(* IEC 61131-3 sources: JingjiangArm/moonboxpro_arm_8.4/Application/Application/任务列表/TensionTask/电机运动/MotionCtl_Gear, 17 files *)

(* ---- StMotorParam_Vel.st ---- *)
(*@CES
Name=StMotorParam_Vel
Type=Gvl
TypeGuid=2db5746d-d284-4425-9f7f-2663a34b0ebc
Guid=35fd48d6-a97b-4a50-89b7-bfdefdaf1e25
HasDeclaration=True
HasImplementation=False
*)
{DECLARATION}
TYPE StMotorParam_Vel :(*速度运动同步轴就是这些各参数了*)
STRUCT
	iAxisId: INT;
	iCoreId: INT;
	iStationId: INT;
	iMoveStep: INT;
	iMotionMode: INT;(*运动模式-=0：电子齿轮=1：JOG=2：点位*)
	xMoveRev: BOOL;
	xMoveEn: BOOL;
	rAxisGirth: REAL;(*同步版周*)
	xMoveVelMode: BOOL;(*=0:线速度=1转速*)
	rAxisVel: REAL;(*速度*)
	uiAxisNum: UINT;(*减速比分子*)
	uiAxisDen: UINT;(*减速比分母*)
	liTargetPos: LINT;(*点位目标位置*)
	udiTargetVel: UDINT;

	//2026.01.31.130843 | + | 增加停机维持伺服功能 秦华有停机维持伺服的功能，需要增加一个判断是否是使能状态的标志
	xAxisOn_ing : BOOL;//此标志表示该轴正处于使能中。。。

	//2026.05.09.085650 | + | 将大指令写入的值先放在这里，然后再穿进去
	modify_delta: DINT;
	/// 可以为正值
	ratio_a: DINT;
	/// 必须为正值
	ratio_b: DINT;

	//2026.05.12.201038 | + | 增加轴单运行中的标志
	xAxisInching : BOOL;
END_STRUCT
END_TYPE

{IMPLEMENTATION}

(* ---- KS_SetMotionCheckServoOn.st ---- *)
(*@CES
Name=KS_SetMotionCheckServoOn
Type=FunctionBlock
TypeGuid=6f9dac99-8de1-4efc-8465-68ac443b7d08
Guid=16f739cf-935e-4f65-a185-0fbe09498330
HasDeclaration=True
HasImplementation=True
*)
{DECLARATION}
FUNCTION KS_SetMotionCheckServoOn : INT
VAR_INPUT
	i_iAxisId: INT;
	i_iCoreId: INT;
	i_iStationId: INT;
	i_pxMoveEn : POINTER TO BOOL;
	i_dwMotionSts: DWORD;
	i_dwDriverSts: DWORD;
	i_pxServoOn: POINTER TO BOOL;
	i_pstStHYLogFifo			: POINTER TO StHYLogFifo;(* 2025.8.23.170701/han.dp/增加的日志队列 *)
END_VAR
VAR
	iResult: INT;
	xRtn: BOOL;
	iFailedAxisCntNum: INT;
	wLogLevel: WORD;
	sMsg_major: STRING;
	sMsg_minor: STRING;
END_VAR

{IMPLEMENTATION}
iResult:= 0;
sMsg_major:= ''; (* 2021.2.26.170203/ *)
sMsg_minor:= ''; (* 2021.2.26.170203/ *)
IF i_iStationId>=1 AND i_iStationId<=MAX_STATION_NUM AND
	i_iAxisId>=1 AND i_iAxisId<=MAX_STATION_NUM AND
	(i_iCoreId=1 OR i_iCoreId=2) THEN

	IF i_pxServoOn^ AND i_pxMoveEn^ THEN
		xRtn:= (*i_dwDriverSts.1 AND*) i_dwMotionSts.9;

		IF NOT xRtn THEN
			iResult:= iResult+1;
			(* 2021.2.26.172210/归属于普通报警 *)
			wLogLevel:= LOG_LEVEL_ALARM_NORMAL;
	(*2022.6.4.093146|精简打印信息！*)
	(*		sMsg_major:= CONCAT('ALARM_NORMAL: KS_SetGrpAxisClrSts_PshLog|Aid:', INT_TO_STRING(iAxisId));*)
			sMsg_major:= CONCAT('KS_SetMotionCheckServoOn|Aid:', INT_TO_STRING(i_iAxisId));
			sMsg_major:= CONCAT(sMsg_major, '|Sid:');
			sMsg_major:= CONCAT(sMsg_major, INT_TO_STRING(i_iStationId));
			sMsg_minor:= CONCAT('CheckServoOn|', BOOL_TO_STRING(xRtn));
			sMsg_minor:= CONCAT(sMsg_minor,'|MotionSts:');
			sMsg_minor:= CONCAT(sMsg_minor, DWORD_TO_STRING(i_dwMotionSts));
		END_IF

		//i_pxServoOn^:= FALSE;
	END_IF
END_IF

IF sMsg_major<>'' THEN (* 2021.2.26.172055/有内容代表要写日志的 *)
	KS_HY_AddMsgToLog(i_pstStHYLogFifo, wLogLevel, sMsg_major, sMsg_minor);
END_IF

KS_SetMotionCheckServoOn:= iResult;

(* ---- KS_SetMotionClrSts.st ---- *)
(*@CES
Name=KS_SetMotionClrSts
Type=FunctionBlock
TypeGuid=6f9dac99-8de1-4efc-8465-68ac443b7d08
Guid=5963aa42-d132-45f6-9961-fbcc83163ad5
HasDeclaration=True
HasImplementation=True
*)
{DECLARATION}
FUNCTION KS_SetMotionClrSts : INT(*0:无错误| >0:失败的指令数量; |-1:参数错误;*)
VAR_INPUT
	i_iAxisId: INT;
	i_iCoreId: INT;
	i_iStationId: INT;
	i_pstStHYLogFifo			: POINTER TO StHYLogFifo;(* 2025.8.23.170701/han.dp/增加的日志队列 *)
END_VAR
VAR
	iResult: INT;
	iRtn: INT;
	iFailedAxisCntNum: INT;
	wLogLevel: WORD;
	sMsg_major: STRING;
	sMsg_minor: STRING;
END_VAR

{IMPLEMENTATION}
iResult:= 0;
sMsg_major:= ''; (* 2021.2.26.170203/ *)
sMsg_minor:= ''; (* 2021.2.26.170203/ *)
IF i_iStationId>=1 AND i_iStationId<=MAX_STATION_NUM AND
	i_iAxisId>=1 AND i_iAxisId<=MAX_STATION_NUM AND
	(i_iCoreId=1 OR i_iCoreId=2) THEN
	iRtn:= GTN_ClrSts(i_iCoreId, i_iAxisId, 1);(*清除错误|*)
	IF iRtn<>0 THEN
		iResult:= iRtn;
		(* 2021.2.26.172210/归属于普通报警 *)
		wLogLevel:= LOG_LEVEL_ALARM;
(*2022.6.4.093146|精简打印信息！*)
(*		sMsg_major:= CONCAT('ALARM_NORMAL: KS_SetGrpAxisClrSts_PshLog|Aid:', INT_TO_STRING(iAxisId));*)
		sMsg_major:= CONCAT('KS_SetMotionClrSts|Aid:', INT_TO_STRING(i_iAxisId));
		sMsg_major:= CONCAT(sMsg_major, '|Sid:');
		sMsg_major:= CONCAT(sMsg_major, INT_TO_STRING(i_iStationId));
		sMsg_minor:= CONCAT('GTN_ClrSts: ', INT_TO_STRING(iRtn));
	END_IF
END_IF

IF sMsg_major<>'' THEN (* 2021.2.26.172055/有内容代表要写日志的 *)
	KS_HY_AddMsgToLog(i_pstStHYLogFifo, wLogLevel, sMsg_major, sMsg_minor);
END_IF

KS_SetMotionClrSts:= iResult;

(* ---- KS_SetMotionMode.st ---- *)
(*@CES
Name=KS_SetMotionMode
Type=FunctionBlock
TypeGuid=6f9dac99-8de1-4efc-8465-68ac443b7d08
Guid=eb1bfde3-c781-4a8b-bb4b-64a6f57a70ed
HasDeclaration=True
HasImplementation=True
*)
{DECLARATION}
FUNCTION KS_SetMotionMode : INT(*0:无错误| >0:失败的指令数量; |-1:参数错误;*)
VAR_INPUT
	i_iAxisId: INT;
	i_iCoreId: INT;
	i_iStationId: INT;
	i_iMoveMode: INT;
	i_iAxisId_Master: INT;
	i_xMasterType : BOOL;
	i_pstStHYLogFifo			: POINTER TO StHYLogFifo;(* 2025.8.23.170701/han.dp/增加的日志队列 *)
END_VAR
VAR
	iResult: INT;
	iRtn: INT;
	iFailedAxisCntNum: INT;
	wLogLevel: WORD;
	sMsg_major: STRING;
	sMsg_minor: STRING;
END_VAR

{IMPLEMENTATION}
iResult:= 0;
sMsg_major:= ''; (* 2021.2.26.170203/ *)
sMsg_minor:= ''; (* 2021.2.26.170203/ *)
IF i_iStationId>=1 AND i_iStationId<=MAX_STATION_NUM AND
	i_iAxisId>=1 AND i_iAxisId<=MAX_STATION_NUM AND
	(i_iCoreId=1 OR i_iCoreId=2) THEN
	IF i_iMoveMode=0 THEN
		iRtn := SetPrfGearModePrm(
				i_iCore:= i_iCoreId,
				i_iAxisId:= i_iAxisId,
				i_iMasterIndex:= i_iAxisId_Master,//i_pastTStGearParamUser^[iCnt_GearAxis].iMasterIndex,
				i_diMasterEven:= 1,//i_pastTStGearParamUser^[iCnt_GearAxis].diMasterEven,
				i_diSlaveEven:= 1,//i_pastTStGearParamUser^[iCnt_GearAxis].diSlaveEven,
				i_diMasterSlope:= 100000,
				i_xMasterType := i_xMasterType);//i_pastTStGearParamUser^[iCnt_GearAxis].diMasterSlope);

	ELSIF i_iMoveMode=1 THEN
		//2025.10.28.105106 | bai.zy  | 单运行仍然使用电子齿轮
		iRtn := SetPrfGearModePrm(
				i_iCore:= i_iCoreId,
				i_iAxisId:= i_iAxisId,
				i_iMasterIndex:= i_iAxisId_Master,//i_pastTStGearParamUser^[iCnt_GearAxis].iMasterIndex,
				i_diMasterEven:= 1,//i_pastTStGearParamUser^[iCnt_GearAxis].diMasterEven,
				i_diSlaveEven:= 1,//i_pastTStGearParamUser^[iCnt_GearAxis].diSlaveEven,
				i_diMasterSlope:= 100000,
				i_xMasterType := i_xMasterType);//i_pastTStGearParamUser^[iCnt_GearAxis].diMasterSlope);

// 		iRtn := SetPrfJogModePrm(
// 				i_iCore:= i_iCoreId,
// 				i_iAxisId:= i_iAxisId,
// 				i_lrAcc:= 1,
// 				i_lrDec:= 1,
// 				i_rSmooth:= 0.8);

	ELSIF i_iMoveMode=2 THEN
		iRtn := SetPrfTrapModePrm(
				i_iCoreId:= i_iCoreId,
				i_iAxisId:= i_iAxisId,
				i_lrVel:= 100,//i_pastTStTrapParamUser^[iCnt_TrapAxis].lrVel,
				i_lrAcc:= 2.0,//i_pastTStTrapParamUser^[iCnt_TrapAxis].lrAcc,
				i_lrDec:= 2.0,//i_pastTStTrapParamUser^[iCnt_TrapAxis].lrDec,
				i_iSmoothTime:= 0);//i_pastTStTrapParamUser^[iCnt_TrapAxis].iSmoothTime);
	ELSIF i_iMoveMode=3 THEN//增加一种运动模式2026.4.27.215724|收放料速度模式
		iRtn := SetPrfJogModePrm(
				i_iCore:= i_iCoreId,
				i_iAxisId:= i_iAxisId,
				i_lrAcc:= 1,
				i_lrDec:= 1,
				i_rSmooth:= 0.8);

	ELSE;
		iRtn := SetPrfGearModePrm(
				i_iCore:= i_iCoreId,
				i_iAxisId:= i_iAxisId,
				i_iMasterIndex:= i_iAxisId_Master,//i_pastTStGearParamUser^[iCnt_GearAxis].iMasterIndex,
				i_diMasterEven:= 1,//i_pastTStGearParamUser^[iCnt_GearAxis].diMasterEven,
				i_diSlaveEven:= 1,//i_pastTStGearParamUser^[iCnt_GearAxis].diSlaveEven,
				i_diMasterSlope:= 100000,
				i_xMasterType := i_xMasterType);//i_pastTStGearParamUser^[iCnt_GearAxis].diMasterSlope);
	END_IF

	IF iRtn<>0 THEN
		iResult:= iRtn;
		(* 2021.2.26.172210/归属于普通报警 *)
		wLogLevel:= LOG_LEVEL_ALARM;
(*2022.6.4.093146|精简打印信息！*)
(*		sMsg_major:= CONCAT('ALARM_NORMAL: KS_SetGrpAxisClrSts_PshLog|Aid:', INT_TO_STRING(iAxisId));*)
		sMsg_major:= CONCAT('KS_SetMotionMode|Aid:', INT_TO_STRING(i_iAxisId));
		sMsg_major:= CONCAT(sMsg_major, '|Sid:');
		sMsg_major:= CONCAT(sMsg_major, INT_TO_STRING(i_iStationId));
		//sMsg_minor:= CONCAT('GTN_ClrSts: ', INT_TO_STRING(iRtn));
	END_IF
END_IF

IF sMsg_major<>'' THEN (* 2021.2.26.172055/有内容代表要写日志的 *)
	KS_HY_AddMsgToLog(i_pstStHYLogFifo, wLogLevel, sMsg_major, sMsg_minor);
END_IF

KS_SetMotionMode:= iResult;

(* ---- KS_SetMotionServoOff.st ---- *)
(*@CES
Name=KS_SetMotionServoOff
Type=FunctionBlock
TypeGuid=6f9dac99-8de1-4efc-8465-68ac443b7d08
Guid=af78d755-d488-4f6e-8233-0470695debbc
HasDeclaration=True
HasImplementation=True
*)
{DECLARATION}
FUNCTION KS_SetMotionServoOff : INT(*0:无错误| >0:失败的指令数量; |-1:参数错误;*)
VAR_INPUT
	i_iAxisId: INT;
	i_iCoreId: INT;
	i_iStationId: INT;
	i_xForceAxisOff:BOOL;(*强制下伺服标志|有效后直接调用AXISOFF指令|2021.5.8.161449*)
	i_dwMotionSts: DWORD;
	i_dwDriverSts: DWORD;
	i_pxServoOn: POINTER TO BOOL;
	i_pstStHYLogFifo			: POINTER TO StHYLogFifo;(* 2025.8.23.170701/han.dp/增加的日志队列 *)
END_VAR
VAR
	iResult: INT;
	iRtn: INT;
	iFailedAxisCntNum: INT;
	wLogLevel: WORD;
	sMsg_major: STRING;
	sMsg_minor: STRING;
END_VAR

{IMPLEMENTATION}
iResult:= 0;
sMsg_major:= ''; (* 2021.2.26.170203/ *)
sMsg_minor:= ''; (* 2021.2.26.170203/ *)
IF i_iStationId>=1 AND i_iStationId<=MAX_STATION_NUM AND
	i_iAxisId>=1 AND i_iAxisId<=MAX_STATION_NUM AND
	(i_iCoreId=1 OR i_iCoreId=2) THEN

	IF i_pxServoOn^ (*OR i_dwDriverSts.1*) THEN
		IF i_xForceAxisOff THEN
			iRtn:= GTN_AxisOff(i_iCoreId, i_iAxisId);
		ELSE
			IF i_dwMotionSts.9=1 THEN
				iRtn:= GTN_AxisOff(i_iCoreId, i_iAxisId);
			ELSE
				iRtn:= 0;
				iResult:= iResult+1;
			END_IF
		END_IF
		IF iRtn<>0 THEN
			iResult:= iResult+1;
			(* 2021.2.26.172210/归属于普通报警 *)
			wLogLevel:= LOG_LEVEL_ALARM;
	(*2022.6.4.093146|精简打印信息！*)
	(*		sMsg_major:= CONCAT('ALARM_NORMAL: KS_SetGrpAxisClrSts_PshLog|Aid:', INT_TO_STRING(iAxisId));*)
			sMsg_major:= CONCAT('KS_SetMotionServoOff|Aid:', INT_TO_STRING(i_iAxisId));
			sMsg_major:= CONCAT(sMsg_major, '|Sid:');
			sMsg_major:= CONCAT(sMsg_major, INT_TO_STRING(i_iStationId));
			sMsg_minor:= CONCAT('GTN_AxisOff: ', INT_TO_STRING(iRtn));
		END_IF
		i_pxServoOn^:= FALSE;
	END_IF
END_IF

IF sMsg_major<>'' THEN (* 2021.2.26.172055/有内容代表要写日志的 *)
	KS_HY_AddMsgToLog(i_pstStHYLogFifo, wLogLevel, sMsg_major, sMsg_minor);
END_IF

KS_SetMotionServoOff:= iResult;

(* ---- KS_SetMotionServoOn.st ---- *)
(*@CES
Name=KS_SetMotionServoOn
Type=FunctionBlock
TypeGuid=6f9dac99-8de1-4efc-8465-68ac443b7d08
Guid=110bff78-641d-4d88-8fec-48f0af46562f
HasDeclaration=True
HasImplementation=True
*)
{DECLARATION}
FUNCTION KS_SetMotionServoOn : INT(*0:无错误| >0:失败的指令数量; |-1:参数错误;*)
VAR_INPUT
	i_iAxisId: INT;
	i_iCoreId: INT;
	i_iStationId: INT;
	i_pxMoveEn : POINTER TO BOOL;
	i_pxServoOn: POINTER TO BOOL;
	i_pstStHYLogFifo			: POINTER TO StHYLogFifo;(* 2025.8.23.170701/han.dp/增加的日志队列 *)
END_VAR
VAR
	iResult: INT;
	iRtn: INT;
	iFailedAxisCntNum: INT;
	wLogLevel: WORD;
	sMsg_major: STRING;
	sMsg_minor: STRING;
END_VAR

{IMPLEMENTATION}
iResult:= 0;
sMsg_major:= ''; (* 2021.2.26.170203/ *)
sMsg_minor:= ''; (* 2021.2.26.170203/ *)
IF i_iStationId>=1 AND i_iStationId<=MAX_STATION_NUM AND
	i_iAxisId>=1 AND i_iAxisId<=MAX_STATION_NUM AND
	(i_iCoreId=1 OR i_iCoreId=2) THEN
	IF i_pxServoOn^ THEN(*如果之前伺服标志被置了,这里先让下伺服|*)
		i_pxServoOn^:= FALSE;
		iRtn := GTN_AxisOff(i_iCoreId, i_iAxisId);
	END_IF

	//2025.10.27.150339 | bai.zy |
	IF i_pxMoveEn^ THEN
		iRtn:= GTN_AxisOn(i_iCoreId, i_iAxisId);(*上伺服|*)
	END_IF

	IF iRtn<>0 THEN
		iResult:= iRtn;
		(* 2021.2.26.172210/归属于普通报警 *)
		wLogLevel:= LOG_LEVEL_ALARM;
(*2022.6.4.093146|精简打印信息！*)
(*		sMsg_major:= CONCAT('ALARM_NORMAL: KS_SetGrpAxisClrSts_PshLog|Aid:', INT_TO_STRING(iAxisId));*)
		sMsg_major:= CONCAT('KS_SetMotionServoOn|Aid:', INT_TO_STRING(i_iAxisId));
		sMsg_major:= CONCAT(sMsg_major, '|Sid:');
		sMsg_major:= CONCAT(sMsg_major, INT_TO_STRING(i_iStationId));
		sMsg_minor:= CONCAT('GTN_AxisOn: ', INT_TO_STRING(iRtn));
		//2026.1.14.200337 | 临时增加 | 观察上伺服失败是什么原因
		iRtn := GTN_AxisOff(i_iCoreId, i_iAxisId);
		iRtn := GTN_ClrSts(i_iCoreId, i_iAxisId, 1);(*清除错误|*)
	ELSE
		IF i_pxMoveEn^ THEN
			i_pxServoOn^:= TRUE;
		END_IF
	END_IF
END_IF

IF sMsg_major<>'' THEN (* 2021.2.26.172055/有内容代表要写日志的 *)
	KS_HY_AddMsgToLog(i_pstStHYLogFifo, wLogLevel, sMsg_major, sMsg_minor);
END_IF

KS_SetMotionServoOn:= iResult;

(* ---- KS_SetMotionZeroPos.st ---- *)
(*@CES
Name=KS_SetMotionZeroPos
Type=FunctionBlock
TypeGuid=6f9dac99-8de1-4efc-8465-68ac443b7d08
Guid=26ac65f6-244c-4574-99d7-e822b9256998
HasDeclaration=True
HasImplementation=True
*)
{DECLARATION}
FUNCTION KS_SetMotionZeroPos : INT
VAR_INPUT
	i_iAxisId: INT;
	i_iCoreId: INT;
	i_iStationId: INT;
	i_pstStHYLogFifo			: POINTER TO StHYLogFifo;(* 2025.8.23.170701/han.dp/增加的日志队列 *)
END_VAR
VAR
	iN: INT;
	iRtn: INT;
	iResult: INT;
	wLogLevel: WORD;
	sMsg_major: STRING;
	sMsg_minor: STRING;
END_VAR

{IMPLEMENTATION}
iResult:= 0;
sMsg_major:= ''; (* 2021.2.26.170203/ *)
sMsg_minor:= ''; (* 2021.2.26.170203/ *)
IF i_iStationId>=1 AND i_iStationId<=MAX_STATION_NUM AND
	i_iAxisId>=1 AND i_iAxisId<=MAX_STATION_NUM AND
	(i_iCoreId=1 OR i_iCoreId=2) THEN
	iRtn:= GTN_ZeroPos(i_iCoreId, i_iAxisId, 1);(*清除错误|*)
	IF iRtn<>0 THEN
		iResult:= iRtn;
		(* 2021.2.26.172210/归属于普通报警 *)
		wLogLevel:= LOG_LEVEL_ALARM;
(*2022.6.4.093146|精简打印信息！*)
(*		sMsg_major:= CONCAT('ALARM_NORMAL: KS_SetGrpAxisClrSts_PshLog|Aid:', INT_TO_STRING(iAxisId));*)
		sMsg_major:= CONCAT('KS_SetMotionZeroPos|Aid:', INT_TO_STRING(i_iAxisId));
		sMsg_major:= CONCAT(sMsg_major, '|Sid:');
		sMsg_major:= CONCAT(sMsg_major, INT_TO_STRING(i_iStationId));
		sMsg_minor:= CONCAT('GTN_ZeroPos: ', INT_TO_STRING(iRtn));
	END_IF
END_IF

IF sMsg_major<>'' THEN (* 2021.2.26.172055/有内容代表要写日志的 *)
	KS_HY_AddMsgToLog(i_pstStHYLogFifo, wLogLevel, sMsg_major, sMsg_minor);
END_IF
KS_SetMotionZeroPos:= iResult;

(* ---- KS_FB_AxisEnCtl.st ---- *)
(*@CES
Name=KS_FB_AxisEnCtl
Type=FunctionBlock
TypeGuid=6f9dac99-8de1-4efc-8465-68ac443b7d08
Guid=7961db84-caed-4243-9b52-56f0bd4c7e60
HasDeclaration=True
HasImplementation=True
*)
{DECLARATION}
FUNCTION_BLOCK KS_FB_AxisEnCtl
VAR_INPUT
	i_xEn: BOOL;
	i_iGrpId: INT;
	i_iGrpUnitNum_Pu : INT;
	i_aiGrpUnitList: ARRAY [1..MAX_UNIT_NUM] OF INT;
	i_iGrpGearMotion_Num: INT;
	i_aiGrpGearMotion_StdList: ARRAY [1..MAX_STATION_NUM] OF INT;
	i_pstStSysParam: POINTER TO StSysParam;
	i_pastStAxisIdListInf :POINTER TO ARRAY [1..128] OF StAxisIdListInf;
	i_pastStMotorParam_Vel: POINTER TO ARRAY [1..MAX_STATION_NUM] OF StMotorParam_Vel;
	i_pstStSysStationInf			:POINTER TO StSysStationInf;
END_VAR
VAR_OUTPUT
	o_iAxisId_Master: INT;
END_VAR
VAR
	iN: INT;
	iAxisId: INT;
	iTypeId: INT;
	iUnitId: INT;
	iCoreId: INT;
	iGroupId : INT;
	pstStGrpParam_Save: POINTER TO StGrpParam_Save;
	pstStGrpParam_UnSave: POINTER TO StGrpParam_UnSave;

	iAdjAxisId : INT;
END_VAR

{IMPLEMENTATION}
IF i_xEn THEN
	IF (i_iGrpId=1 OR i_iGrpId=2) AND
		i_iGrpUnitNum_Pu>=1 AND i_iGrpUnitNum_Pu<=MAX_UNIT_NUM AND
		i_iGrpGearMotion_Num>=1 AND i_iGrpGearMotion_Num<= MAX_STATION_NUM AND
		i_pstStSysParam<>0 AND
		i_pastStAxisIdListInf<>0 AND
		i_pastStMotorParam_Vel<>0 AND
		i_pstStSysStationInf <> 0 THEN
		pstStGrpParam_Save:= ADR(i_pstStSysParam^.astStGrpParam_Save[i_iGrpId]);
		pstStGrpParam_UnSave:= ADR(i_pstStSysParam^.astStGrpParam_UnSave[i_iGrpId]);

		FOR iN:=1 TO i_iGrpGearMotion_Num BY 1 DO
// 			KS_HY_GetAxisIdForMotByStation(
// 				i_aiGrpGearMotion_StdList[iN],
// 				ADR(iAxisId),
// 				ADR(iTypeId),
// 				ADR(iUnitId),
// 				ADR(iCoreId),
// 				ADR(iGroupId),
// 				ADR(iAdjAxisId),
// 				i_pastStAxisIdListInf);
			KS_GetAxisIdForMotByStation_V2(
					i_iStationId:= i_aiGrpGearMotion_StdList[iN],
					i_piAxisId:= ADR(iAxisId),
					i_piTypeId:= ADR(iTypeId),
					i_piUnitId:= ADR(iUnitId),
					i_piCoreId:= ADR(iCoreId),
					i_piGroupId:= ADR(iGroupId),
					i_piAdjAxisId:= ADR(iAdjAxisId),
					i_pstStSysStationInf:= i_pstStSysStationInf);
			CASE iTypeId OF
			TYPE_MASTER_I,TYPE_MASTER_II:
				o_iAxisId_Master:= iAxisId;
			TYPE_CENTRAL_I,TYPE_CENTRAL_II:
				i_pastStMotorParam_Vel^[iN].xMoveEn:= pstStGrpParam_UnSave^.xFlag_Print;
				i_pastStMotorParam_Vel^[iN].xMoveRev:= pstStGrpParam_UnSave^.xMotRev_CentralDrum;
				i_pastStMotorParam_Vel^[iN].xMoveVelMode:= TRUE;
			TYPE_UNWIND_A_I,TYPE_UNWIND_A_II:
				i_pastStMotorParam_Vel^[iN].xMoveEn:= pstStGrpParam_UnSave^.xAxisAForeward_Uw;
				i_pastStMotorParam_Vel^[iN].xMoveRev:= pstStGrpParam_UnSave^.xMotRev_AxisA_Uw;
				i_pastStMotorParam_Vel^[iN].xMoveVelMode:= FALSE;
			TYPE_UNWIND_B_I,TYPE_UNWIND_B_II:
				i_pastStMotorParam_Vel^[iN].xMoveEn:= pstStGrpParam_UnSave^.xAxisBForeward_Uw;
				i_pastStMotorParam_Vel^[iN].xMoveRev:= pstStGrpParam_UnSave^.xMotRev_AxisB_Uw;
				i_pastStMotorParam_Vel^[iN].xMoveVelMode:= FALSE;
			TYPE_REWIND_A_I,TYPE_REWIND_A_II:
				i_pastStMotorParam_Vel^[iN].xMoveEn:= pstStGrpParam_UnSave^.xAxisAForeward_Rw;
				i_pastStMotorParam_Vel^[iN].xMoveRev:= pstStGrpParam_UnSave^.xMotRev_AxisA_Rw;
				i_pastStMotorParam_Vel^[iN].xMoveVelMode:= FALSE;
			TYPE_REWIND_B_I,TYPE_REWIND_B_II:
				i_pastStMotorParam_Vel^[iN].xMoveEn:= pstStGrpParam_UnSave^.xAxisBForeward_Rw;
				i_pastStMotorParam_Vel^[iN].xMoveRev:= pstStGrpParam_UnSave^.xMotRev_AxisB_Rw;
				i_pastStMotorParam_Vel^[iN].xMoveVelMode:= FALSE;
			TYPE_INFEED_I,TYPE_INFEED_II:
				i_pastStMotorParam_Vel^[iN].xMoveEn:= pstStGrpParam_UnSave^.xFlag_Print OR pstStGrpParam_UnSave^.xFlag_Ink OR i_pstStSysParam^.astStRSV_GrpParam_UnSave[i_iGrpId].xInching_If_Roller;
				i_pastStMotorParam_Vel^[iN].xMoveRev:= pstStGrpParam_UnSave^.xMotRev_If;
				i_pastStMotorParam_Vel^[iN].xMoveVelMode:= TRUE;
			TYPE_OUTFEED_I,TYPE_OUTFEED_II:
				i_pastStMotorParam_Vel^[iN].xMoveEn:= pstStGrpParam_UnSave^.xFlag_Print OR pstStGrpParam_UnSave^.xFlag_Ink OR i_pstStSysParam^.astStRSV_GrpParam_UnSave[i_iGrpId].xInching_Of_Roller;
				i_pastStMotorParam_Vel^[iN].xMoveRev:= pstStGrpParam_UnSave^.xMotRev_Of;
				i_pastStMotorParam_Vel^[iN].xMoveVelMode:= TRUE;
			TYPE_UNIT_PRN:
				i_pastStMotorParam_Vel^[iN].xMoveEn:= i_pstStSysParam^.astStUnitParam_UnSave[iUnitId].xEn_Motor_PrnRoller;
				i_pastStMotorParam_Vel^[iN].xMoveRev:= i_pstStSysParam^.astStUnitParam_UnSave[iUnitId].xMotRev_PrnRoller;
				i_pastStMotorParam_Vel^[iN].xMoveVelMode:= TRUE;
			TYPE_UNIT_BOTTOM:
				i_pastStMotorParam_Vel^[iN].xMoveEn:= i_pstStSysParam^.astStUnitParam_UnSave[iUnitId].xEn_Motor_BottomRoller;
				i_pastStMotorParam_Vel^[iN].xMoveRev:= i_pstStSysParam^.astStUnitParam_UnSave[iUnitId].xMotRev_BottomRoller;
				i_pastStMotorParam_Vel^[iN].xMoveVelMode:= TRUE;
			TYPE_UNIT_NET:
				i_pastStMotorParam_Vel^[iN].xMoveEn:= i_pstStSysParam^.astStUnitParam_UnSave[iUnitId].xEn_Motor_NetRoller;
				i_pastStMotorParam_Vel^[iN].xMoveRev:= i_pstStSysParam^.astStUnitParam_UnSave[iUnitId].xMotRev_NetRoller;
				i_pastStMotorParam_Vel^[iN].xMoveVelMode:= TRUE;
			END_CASE
		END_FOR
	END_IF
ELSE
	;
END_IF

(* ---- KS_FB_AxisInchCtl.st ---- *)
(*@CES
Name=KS_FB_AxisInchCtl
Type=FunctionBlock
TypeGuid=6f9dac99-8de1-4efc-8465-68ac443b7d08
Guid=962c4a2d-5100-4818-8083-96730c4559b1
HasDeclaration=True
HasImplementation=True
*)
{DECLARATION}
FUNCTION_BLOCK KS_FB_AxisInchCtl
VAR_INPUT
	i_xEn: BOOL;(*使能|*)
	i_iGrpId: INT;(*系id|*)
	i_iGrpAxisNum_Pu: INT;(*色组轴的数量|*)
	i_aiGrpAxisList: ARRAY [1..MAX_UNIT_NUM] OF INT;(*系内所有轴的id列表,色组部分已经按照从小到大的顺序排序了，之后的是牵引|*)
	i_pstStSysParam: POINTER TO StSysParam;(*参数结构|*)
//	i_pastStPTSts: POINTER TO ARRAY [1..MAX_STATION_NUM] OF StPTSts;(*PT运动轴的状态|*)
	i_pastStIOMap_Main_FE						: POINTER TO ARRAY [1..4] OF StIOMap_Main_FE;(*轴io数据区域|AB系*)
	i_pastStIOMap_Axis_FE					: POINTER TO ARRAY [1..MAX_UNIT_NUM] OF StIOMap_Axis_FE;(*轴io数据区域|`````````````````````````````````````````````*)
	i_pstStEvtReq: POINTER TO StEvtReq;(*输入动作|*)
	i_xAllLinkageAxis_Inch:BOOL;(*2022.5.21.103459 所有联动轴单运行功能使能标志*)
END_VAR
VAR_OUTPUT
	o_xEno: BOOL;(*Same with i_xEn|*)
	o_iErNo: INT;(*-1参数错误\|*)
	o_xHasAxisOnInchRunningSts: BOOL;(*True标识有轴还在单运行|*)
	o_diVel_Virtual_Tar_Inch: DINT;(*虚拟主轴规划速度*)
	o_lrMax_a_S_pos_Inch: LREAL;(*虚拟主轴最大减速度*)
	o_arInchTarVel : ARRAY [1..MAX_UNIT_NUM] OF REAL;
END_VAR
VAR
	iN: INT;
	iUnitId: INT;
	pstStGrpParam_Save: POINTER TO StGrpParam_Save;
	pstStGrpParam_UnSave: POINTER TO StGrpParam_UnSave;
	pstStUnitParam_Save: POINTER TO StUnitParam_Save;
	pstStUnitParam_UnSave: POINTER TO StUnitParam_UnSave;
	axAxisInching_Temp:ARRAY [1..MAX_UNIT_NUM] OF BOOL;(*轴单运行中@无效的时候不一定是真正的0速*)
	axInchPressReq: ARRAY [1..MAX_UNIT_NUM] OF BOOL := [MAX_UNIT_NUM(FALSE)];
	pstStIOMap_Axis_FE					: POINTER TO StIOMap_Axis_FE;(*轴io数据区域|`````````````````````````````````````````````*)
	abyAxisMoveSts:ARRAY [1..MAX_UNIT_NUM] OF BYTE;(*轴运动状态@=1 单运行状态|=2 jog运动状态|=3 等待状态*)
	axInchAxisRev:ARRAY [1..MAX_UNIT_NUM] OF BOOL;(*反转标志处理@默认是正转*)
	axFlag_Inched : ARRAY [1..MAX_UNIT_NUM] OF BOOL := [MAX_UNIT_NUM(FALSE)];
	axAxisInchAutoAccing:ARRAY [1..MAX_STATION_NUM] OF BOOL;(*轴单运行自动加速中*)
	arInchTarVel: ARRAY [1..MAX_STATION_NUM] OF REAL;
	iInchMaxVel:INT:=50;(*单运行最大速度*)
	xAccBtn: BOOL;
	xDecBtn: BOOL;
	lrTmp:LREAL;

	//2025.10.28.140624 | bai.zy | 单运行的轴速度先单独拿出来
	adiVel_Virtual_Tar_Inch : ARRAY [1..MAX_UNIT_NUM] OF DINT;
END_VAR

{IMPLEMENTATION}
(*////////////////////////////////////////*)
(*2019.6.14.092753|单运行增加整机单运行|联动色组按下单运行后所有联动色进入单运行*)
(*////////////////////////////////////////*)
o_xEno:= i_xEn;
o_iErNo:= 0;(*初始化错误代码|*)
o_xHasAxisOnInchRunningSts:= FALSE;
IF i_xEn THEN
	IF (i_iGrpId=1 OR i_iGrpId=2) AND
		(i_iGrpAxisNum_Pu>=1 AND i_iGrpAxisNum_Pu<=MAX_STATION_NUM) AND
		i_pstStSysParam<>0 AND

		i_pastStIOMap_Main_FE<>0 AND
		i_pastStIOMap_Axis_FE<>0 AND
		i_pstStEvtReq<>0 THEN(*2019.6.13.191036|*)
		(*the parameters are valid|*)
		pstStGrpParam_Save:= ADR(i_pstStSysParam^.astStGrpParam_Save[i_iGrpId]);
		pstStGrpParam_UnSave:= ADR(i_pstStSysParam^.astStGrpParam_UnSave[i_iGrpId]);
		(*2022.5.21.103542*)
		IF i_xAllLinkageAxis_Inch THEN;
		ELSE(*不允许整机单运行|*)
			i_pstStEvtReq^.xReqAllInchRun:=FALSE;(*屏蔽按钮*)
		END_IF

		IF i_pstStSysParam^.stStSysParam_Save.xWorkMode_Inch THEN(*单运行方式true一次走一次停*)
			(*先识别动作|*)
			(*整机|*)
			IF i_pstStEvtReq^.xReqAllInchRun THEN(*按了整机单运行|联动色组的单运行也是作为整机单运行处理||*)
				pstStGrpParam_UnSave^.xFlag_AllInchRun:= NOT pstStGrpParam_UnSave^.xFlag_AllInchRun;(*切换单运行状态|*)
			END_IF
			(*2023.6.18.231611 条件优化*)
(*			FOR iN:=1 TO i_iGrpAxisNum_Pu BY 1 DO*)
			FOR iN:=1 TO i_iGrpAxisNum_Pu BY 1 DO(*条件优化@2023.6.16.132433*)
				iUnitId:= i_aiGrpAxisList[iN];(*轴id|*)
				pstStUnitParam_Save:= ADR(i_pstStSysParam^.astStUnitParam_Save[iUnitId]);
				pstStUnitParam_UnSave:= ADR(i_pstStSysParam^.astStUnitParam_UnSave[iUnitId]);
				IF pstStUnitParam_Save^.xLinkage AND
(*						pstStAxisParam^.xAxisInching<>pstStGrpParam^.xFlag_AllInchRun*)
					axAxisInching_Temp[iUnitId]<>pstStGrpParam_UnSave^.xFlag_AllInchRun THEN
(*						pstStAxisParam^.xAxisInching:= pstStGrpParam^.xFlag_AllInchRun;*)
					(*2023.6.18.232053 替换为了临时变量*)
					axAxisInching_Temp[iUnitId]:= pstStGrpParam_UnSave^.xFlag_AllInchRun;
				END_IF

			END_FOR

			(*单动轴|*)
			FOR iN:=1 TO i_iGrpAxisNum_Pu BY 1 DO
				iUnitId:= i_aiGrpAxisList[iN];(*轴id|*)
				pstStUnitParam_Save:= ADR(i_pstStSysParam^.astStUnitParam_Save[iUnitId]);
				pstStUnitParam_UnSave:= ADR(i_pstStSysParam^.astStUnitParam_UnSave[iUnitId]);
				IF (NOT pstStUnitParam_Save^.xLinkage) AND
					(NOT axInchPressReq[iUnitId]) AND
					axInchPressReq[iUnitId]<>i_pastStIOMap_Axis_FE^[iUnitId].i_xInch THEN
	(*					pstStAxisParam^.xAxisInching:= NOT pstStAxisParam^.xAxisInching;*)
					(*2023.6.18.232053 替换为了临时变量*)
					axAxisInching_Temp[iUnitId]:= NOT axAxisInching_Temp[iUnitId];
				END_IF
			END_FOR
		ELSE(*按住走松开停*)
		(*整机|*)
			pstStGrpParam_UnSave^.xFlag_AllInchRun:=i_pstStEvtReq^.xEvt_AllInchRun;(*切换当运行状态*)
			(*条件优化@2023.6.18.231700*)
(*			FOR iN:=1 TO i_iGrpAxisNum_Pu BY 1 DO*)
			FOR iN:=1 TO i_iGrpAxisNum_Pu BY 1 DO
				iUnitId:= i_aiGrpAxisList[iN];(*轴id|*)
				pstStUnitParam_Save:= ADR(i_pstStSysParam^.astStUnitParam_Save[iUnitId]);
				pstStUnitParam_UnSave:= ADR(i_pstStSysParam^.astStUnitParam_UnSave[iUnitId]);
(*					pstStAxisParam^.xAxisInching:= pstStGrpParam^.xFlag_AllInchRun
													AND pstStAxisParam^.xLinkage;(*2019.12.6.110501|增加了联动条件|Liu.yt*)*)
					(*2023.6.18.232053 替换为了临时变量*)
				axAxisInching_Temp[iUnitId]:= pstStGrpParam_UnSave^.xFlag_AllInchRun
													AND pstStUnitParam_Save^.xLinkage;(*2019.12.6.110501|增加了联动条件|Liu.yt*)

			END_FOR

			(*单动轴|*)
			FOR iN:=1 TO i_iGrpAxisNum_Pu BY 1 DO
				iUnitId:= i_aiGrpAxisList[iN];(*轴id|*)
				pstStUnitParam_Save:= ADR(i_pstStSysParam^.astStUnitParam_Save[iUnitId]);
				pstStUnitParam_UnSave:= ADR(i_pstStSysParam^.astStUnitParam_UnSave[iUnitId]);
				IF (NOT pstStUnitParam_Save^.xLinkage) THEN
(*					pstStAxisParam^.xAxisInching:= axInchPressReq[iAxisId];*)
					(*2023.6.18.232053 替换为了临时变量*)
					axAxisInching_Temp[iUnitId]:=axInchPressReq[iUnitId];
				END_IF
			END_FOR
		END_IF

(*2025.10.23.160344这里先放着后面细看处理start*)
		(*兼容单运行和jog模式*)
		FOR iN:=1 TO i_iGrpAxisNum_Pu BY 1 DO
			iUnitId:= i_aiGrpAxisList[iN];(*轴id|*)
			pstStUnitParam_Save:= ADR(i_pstStSysParam^.astStUnitParam_Save[iUnitId]);
			pstStUnitParam_UnSave:= ADR(i_pstStSysParam^.astStUnitParam_UnSave[iUnitId]);
			pstStIOMap_Axis_FE:=ADR(i_pastStIOMap_Axis_FE^[iUnitId]);
			CASE abyAxisMoveSts[iUnitId] OF
				1:(*单运行状态*)
					pstStUnitParam_UnSave^.xAxisInching:= axAxisInching_Temp[iUnitId];
					axInchAxisRev[iUnitId]:= FALSE;//i_pstStShmGlobalParam^.astStGrpParam[i_iGrpId].xUnitRev;(*方向控制*)
					IF NOT pstStUnitParam_UnSave^.xAxisInching AND(*退出了单运行*)
						NOT g_axAxisInching[iUnitId] (*AND(*完全退出了单运行*)		//2025.10.28.114601 | bai.zy | 屏蔽状态机
						pstStAxisParam^.iAxisInchingCaseId=MOTION_STEP_Nothing*) THEN(*退出到初始状态了*)
						abyAxisMoveSts[iUnitId]:=0;
					END_IF
				2:(*JOG状态*)
					IF (NOT pstStUnitParam_Save^.xLinkage) THEN
						pstStUnitParam_UnSave^.xAxisInching:=axAxisInching_Temp[iUnitId];
								(*pstStIOMap_AxisBasic^.i_xServoJog_For OR		//2025.10.28.114601 | bai.zy | 屏蔽方向
								pstStIOMap_AxisBasic^.i_xServoJog_Rev;
						IF pstStIOMap_AxisBasic^.i_xServoJog_Rev THEN
							axInchAxisRev[iUnitId]:=TRUE;(*方向控制*)
						ELSIF pstStIOMap_AxisBasic^.i_xServoJog_For THEN
							axInchAxisRev[iUnitId]:=FALSE;(*方向控制*)
						ELSE(*完全停止了*)
							abyAxisMoveSts[iUnitId]:=3;
						END_IF
						*)
						IF NOT pstStUnitParam_UnSave^.xAxisInching THEN
							abyAxisMoveSts[iUnitId]:=3;
						END_IF
					ELSE(*联动了@清除标志退出case*)
						pstStUnitParam_UnSave^.xAxisInching:=FALSE;
						abyAxisMoveSts[iUnitId]:=3;
					END_IF

				3:(*等待状态*)
					IF NOT pstStUnitParam_UnSave^.xAxisInching AND(*退出了单运行*)
						NOT g_axAxisInching[iUnitId] (*AND(*完全退出了单运行*)		//2025.10.28.114601 | bai.zy | 屏蔽状态机
						pstStAxisParam^.iAxisInchingCaseId=MOTION_STEP_Nothing*) THEN(*退出到初始状态了*)
						abyAxisMoveSts[iUnitId]:=0;
					END_IF

			ELSE
				(*单运行控制@这里只需要赋值就好*)
				pstStUnitParam_UnSave^.xAxisInching:= axAxisInching_Temp[iUnitId];
				abyAxisMoveSts[iUnitId]:=BOOL_TO_BYTE(pstStUnitParam_UnSave^.xAxisInching);(*2023.6.16.132359*)

				IF (NOT pstStUnitParam_Save^.xLinkage) THEN
					(*jog控制@优先单运行*)
					IF NOT pstStUnitParam_UnSave^.xAxisInching THEN
						pstStUnitParam_UnSave^.xAxisInching:=axAxisInching_Temp[iUnitId];
								(*pstStIOMap_AxisBasic^.i_xServoJog_For OR		//2025.10.28.114601 | bai.zy | 屏蔽方向
								pstStIOMap_AxisBasic^.i_xServoJog_Rev;*)
						IF pstStUnitParam_UnSave^.xAxisInching THEN
							abyAxisMoveSts[iUnitId]:=2;
						END_IF
					END_IF
				END_IF
			END_CASE
		END_FOR
(*2025.10.23.160344这里先放着后面细看处理end*)

		IF NOT pstStGrpParam_UnSave^.xFlag_Stop OR (*非停机状态下,禁止各种形式的单运行*)
			(i_pstStEvtReq^.xReqStop AND pstStGrpParam_UnSave^.xFlag_Stop) THEN(*2021.10.15.094231 增加按下停止按钮时候清除单运行*)
			FOR iN:=1 TO i_iGrpAxisNum_Pu BY 1 DO
				iUnitId:= i_aiGrpAxisList[iN];(*轴id|*)
				pstStUnitParam_Save:= ADR(i_pstStSysParam^.astStUnitParam_Save[iUnitId]);
				pstStUnitParam_UnSave:= ADR(i_pstStSysParam^.astStUnitParam_UnSave[iUnitId]);
				pstStUnitParam_UnSave^.xAxisInching:=FALSE;
				axAxisInching_Temp[iUnitId]:=FALSE;(*2023.6.18.232805@无效的时候不一定是真正的0速*)
				abyAxisMoveSts[iUnitId]:=0;(*2023.6.18.231830*)
			END_FOR
			(*非停机的时候清除全体运行标志|2019.12.6.110407*)
			pstStGrpParam_UnSave^.xFlag_AllInchRun:=FALSE;
		END_IF

		(*2025.1.13.182252+*)
		IF pstStGrpParam_UnSave^.xFlag_Home OR
			pstStGrpParam_UnSave^.xFlag_PreRegister OR
			pstStGrpParam_UnSave^.xFlag_PhaseRestore OR
			pstStGrpParam_UnSave^.xFlag_PhaseRead THEN
			pstStGrpParam_UnSave^.xFlag_AllInchRun:=FALSE;
		END_IF
		(*移位到aaaa处|2020.10.12.161828*)

	ELSE
		o_iErNo:= -1;(*参数非法|*)
	END_IF
ELSE
	IF (i_iGrpId=1 OR i_iGrpId=2) AND
		(i_iGrpAxisNum_Pu>=1 AND i_iGrpAxisNum_Pu<=MAX_STATION_NUM) AND
		i_pstStSysParam<>0 AND

		i_pastStIOMap_Main_FE<>0 AND
		i_pastStIOMap_Axis_FE<>0 AND
		i_pstStEvtReq<>0 THEN(*2019.6.13.191036|*)
		(*the parameters are valid|*)

		pstStGrpParam_Save:= ADR(i_pstStSysParam^.astStGrpParam_Save[i_iGrpId]);
		pstStGrpParam_UnSave:= ADR(i_pstStSysParam^.astStGrpParam_UnSave[i_iGrpId]);
		FOR iN:=1 TO i_iGrpAxisNum_Pu BY 1 DO
			iUnitId:= i_aiGrpAxisList[iN];(*轴id|*)
			pstStUnitParam_Save:= ADR(i_pstStSysParam^.astStUnitParam_Save[iUnitId]);
			pstStUnitParam_UnSave:= ADR(i_pstStSysParam^.astStUnitParam_UnSave[iUnitId]);
//			iStationId:= pstStAxisParam^.iStationId;(*站id|*)
			axFlag_Inched[iUnitId]:=FALSE;
			i_pastStIOMap_Axis_FE^[iUnitId].o_xLamp_Inch:= FALSE;
			pstStUnitParam_UnSave^.xAxisInching:=FALSE;
			axAxisInching_Temp[iUnitId]:=FALSE;(*2023.6.18.232805*)
			abyAxisMoveSts[iUnitId]:=0;(*2023.6.18.231830*)
(*
			g_axAxisInchDecing[iAxisId]:=FALSE;
			g_axAxisInching[iAxisId]:=FALSE;*)
		END_FOR
		o_xHasAxisOnInchRunningSts:= FALSE;

		pstStGrpParam_UnSave^.xFlag_AllInchRun:= FALSE; (* 2020.10.12.114752|将整机单运行标志清除掉 *)
	END_IF
END_IF

IF i_pstStSysParam<>0 AND

	i_pastStIOMap_Main_FE<>0 AND
	i_pastStIOMap_Axis_FE<>0 AND
	i_pstStEvtReq<>0 THEN(*2019.6.13.191036|*)
	pstStGrpParam_Save:= ADR(i_pstStSysParam^.astStGrpParam_Save[i_iGrpId]);
	pstStGrpParam_UnSave:= ADR(i_pstStSysParam^.astStGrpParam_UnSave[i_iGrpId]);
	(*aaaa*)
	FOR iN:=1 TO i_iGrpAxisNum_Pu  BY 1 DO
		iUnitId:= i_aiGrpAxisList[iN];(*轴id|*)
		pstStUnitParam_Save:= ADR(i_pstStSysParam^.astStUnitParam_Save[iUnitId]);
		pstStUnitParam_UnSave:= ADR(i_pstStSysParam^.astStUnitParam_UnSave[iUnitId]);
		pstStIOMap_Axis_FE:=ADR(i_pastStIOMap_Axis_FE^[iUnitId]);
	//	iStationId:= pstStAxisParam^.iStationId;(*站id|*)
	//	pstAxisStPTSts:= ADR(i_pastStPTSts^[iAxisId]);(*PTSts|*)

		(*2022.2.15.141220*)
		xAccBtn:=pstStIOMap_Axis_FE^.i_xAcc;
		xDecBtn:=pstStIOMap_Axis_FE^.i_xDec;
		IF pstStGrpParam_UnSave^.xFlag_AllInchRun THEN(*如果是整机点运行|加减速使用整机加减速按钮*)
			xAccBtn:=i_pstStEvtReq^.xEvt_ManuSpdUp;
			xDecBtn:=i_pstStEvtReq^.xEvt_ManuSpdDn;
		END_IF

		(*2019.10.23.155917 对单运行停止做规划,不再像以前一样直接下伺服|Liu.yt---START*)
		IF pstStUnitParam_UnSave^.xAxisInching THEN
			IF NOT g_axAxisInching[iUnitId] THEN(*先自动加速到单运行速度*)
				g_axAxisInching[iUnitId]:=TRUE;
				g_axAxisInchAccing[iUnitId]:=TRUE;
				g_axAxisInchDecing[iUnitId]:=FALSE;
				axAxisInchAutoAccing[iUnitId]:=TRUE;
				arInchTarVel[iUnitId]:= pstStGrpParam_Save^.rVel_Inch;
			END_IF

			IF axAxisInchAutoAccing[iUnitId] THEN
				IF pstStUnitParam_UnSave^.rAxisVel_PrnRoller= pstStGrpParam_Save^.rVel_Inch THEN(*到达目标速度*)
					axAxisInchAutoAccing[iUnitId]:=FALSE;
				END_IF

				IF xAccBtn OR
					xDecBtn THEN
					axAxisInchAutoAccing[iUnitId]:=FALSE;
				END_IF
			ELSE
				g_axAxisInchAccing[iUnitId]:=FALSE;
				g_axAxisInchDecing[iUnitId]:=FALSE;
				IF xAccBtn THEN
					g_axAxisInchAccing[iUnitId]:=TRUE;
					g_axAxisInchDecing[iUnitId]:=FALSE;
					arInchTarVel[iUnitId]:=INT_TO_REAL(iInchMaxVel);(**)
				ELSIF xDecBtn THEN
					g_axAxisInchAccing[iUnitId]:=FALSE;
					g_axAxisInchDecing[iUnitId]:=TRUE;
				END_IF
			END_IF
		ELSIF g_axAxisInching[iUnitId] THEN
			axAxisInchAutoAccing[iUnitId]:=FALSE;
			g_axAxisInchAccing[iUnitId]:=FALSE;
			g_axAxisInchDecing[iUnitId]:=TRUE;
			IF pstStUnitParam_UnSave^.rAxisVel_PrnRoller = 0 THEN
				g_axAxisInchDecing[iUnitId]:=FALSE;
				g_axAxisInching[iUnitId]:=FALSE;
			END_IF
		END_IF
		(*2019.10.23.155917 对单运行停止做规划,不再像以前一样直接下伺服|Liu.yt---END*)
	(*放速度规划吧2025.10.23.164518*)
		IF 	pstStUnitParam_UnSave^.xAxisInching OR g_axAxisInchDecing[iUnitId] THEN
// 			IF pstStUnitParam_UnSave^.iAxisPrnRunCaseId=MOTION_STEP_Nothing THEN(*这里做速度规划-让主轴先动起来*)
// 				//2025.10.28.113117 | bai.zy | 在此处转换成脉冲每毫秒
// 				//o_diVel_Virtual_Tar_Inch:= LREAL_TO_DINT(arInchTarVel[iUnitId]);
// 				o_diVel_Virtual_Tar_Inch:= LREAL_TO_DINT(arInchTarVel[iUnitId]*GC_LRMOTORPPR/pstStUnitParam_Save^.rGirth_PrnRoller/60.0);
// 				o_lrMax_a_S_pos_Inch:= 0.2;
// 			ELSE(*这里规划单运行轴的轴速度*)
				//2025.10.28.113117 | bai.zy | 在此处转换成脉冲每毫秒
				//o_diVel_Virtual_Tar_Inch:= LREAL_TO_DINT(arInchTarVel[iUnitId]);
				//o_diVel_Virtual_Tar_Inch:= LREAL_TO_DINT(arInchTarVel[iUnitId]*GC_LRMOTORPPR/pstStUnitParam_Save^.rGirth_PrnRoller/60.0);
				adiVel_Virtual_Tar_Inch[iUnitId] := LREAL_TO_DINT(arInchTarVel[iUnitId]*GC_LRMOTORPPR/
																gc_rGirth_Master/60.0/1000);
				o_lrMax_a_S_pos_Inch:= 0.2;
				IF g_axAxisInchAccing[iUnitId] THEN
					(*单运行的加速做点处理@在开始的时候加速慢一点,到达一定速度后再加快,方便预套准对mark线*)
					IF ABS(pstStUnitParam_UnSave^.rAxisVel_PrnRoller)>3 THEN
						lrTmp:=0.2;
					ELSE
						lrTmp:=0.04;
					END_IF

					pstStUnitParam_UnSave^.rAxisVel_PrnRoller:= pstStUnitParam_UnSave^.rAxisVel_PrnRoller+lrTmp;(*2025.1.15.150454 调整*)
					IF pstStUnitParam_UnSave^.rAxisVel_PrnRoller>=arInchTarVel[iUnitId] THEN
						pstStUnitParam_UnSave^.rAxisVel_PrnRoller:= arInchTarVel[iUnitId];
					END_IF
				ELSIF g_axAxisInchDecing[iUnitId] THEN(*单运行减速中*)
					pstStUnitParam_UnSave^.rAxisVel_PrnRoller:= pstStUnitParam_UnSave^.rAxisVel_PrnRoller-0.4;(*减速快一点*)
					IF pstStUnitParam_UnSave^.rAxisVel_PrnRoller<=0 THEN
						pstStUnitParam_UnSave^.rAxisVel_PrnRoller:= 0;
					END_IF
				END_IF
				IF NOT o_xHasAxisOnInchRunningSts THEN
					o_xHasAxisOnInchRunningSts:= TRUE;
				END_IF
			//END_IF
		ELSE
			o_xHasAxisOnInchRunningSts:= FALSE;
			//o_diVel_Virtual_Tar_Inch:= 0;
			adiVel_Virtual_Tar_Inch[iUnitId] := 0;
			o_lrMax_a_S_pos_Inch:= 0.2;
		END_IF

	END_FOR

	//2025.10.28.140948 | bai.zy | 输出速度
	FOR iN := 1 TO i_iGrpAxisNum_Pu BY 1 DO
		pstStUnitParam_Save:= ADR(i_pstStSysParam^.astStUnitParam_Save[iN]);
		pstStUnitParam_UnSave:= ADR(i_pstStSysParam^.astStUnitParam_UnSave[iN]);
		IF (pstStUnitParam_UnSave^.xAxisInching OR pstStGrpParam_UnSave^.xFlag_AllInchRun) AND adiVel_Virtual_Tar_Inch[iN] <> 0 THEN
			o_diVel_Virtual_Tar_Inch :=  adiVel_Virtual_Tar_Inch[iN];
			EXIT;
		END_IF
	END_FOR
END_IF

IF i_pastStIOMap_Axis_FE<>0 THEN
	FOR iN:=1 TO MAX_UNIT_NUM BY 1 DO
		axInchPressReq[iN]:= i_pastStIOMap_Axis_FE^[iN].i_xInch;
		o_arInchTarVel[iN] := i_pstStSysParam^.astStUnitParam_UnSave[iN].rAxisVel_PrnRoller;
	END_FOR
END_IF

(* ---- KS_FB_AxisInchCtl_All.st ---- *)
(*@CES
Name=KS_FB_AxisInchCtl_All
Type=FunctionBlock
TypeGuid=6f9dac99-8de1-4efc-8465-68ac443b7d08
Guid=891b7f07-929e-4459-bfed-60e763b2668b
HasDeclaration=True
HasImplementation=True
*)
{DECLARATION}
FUNCTION_BLOCK KS_FB_AxisInchCtl_All
VAR_INPUT
	i_xEn: BOOL;(*使能|*)
	i_iGrpId: INT;(*系id|*)
	i_iGrpAxisNum_Pu: INT;(*色组轴的数量|*)
	i_aiGrpAxisList: ARRAY [1..MAX_UNIT_NUM] OF INT;(*系内所有轴的id列表,色组部分已经按照从小到大的顺序排序了，之后的是牵引|*)
	i_pstStSysParam: POINTER TO StSysParam;(*参数结构|*)
	i_pstStEvtReq: POINTER TO StEvtReq;(*输入动作|*)
	i_pastStIOMap_Axis_FE					: POINTER TO ARRAY [1..MAX_UNIT_NUM] OF StIOMap_Axis_FE;(*轴io数据区域*)
	i_rAcc_Inch : REAL := 0.2;
END_VAR
VAR_OUTPUT
	o_xEno: BOOL;(*Same with i_xEn|*)
	o_iErNo: INT;(*-1参数错误\|*)
	o_xHasAxisOnInchRunningSts: BOOL;(*True标识有轴还在单运行|*)
	o_diVel_Virtual_Tar_Inch: DINT;(*虚拟主轴规划速度*)
	o_lrMax_a_S_pos_Inch: LREAL;(*虚拟主轴最大减速度*)
	o_arInchTarVel : ARRAY [1..MAX_UNIT_NUM] OF REAL;
	o_xInchDecing : BOOL;
END_VAR
VAR
	iN: INT;
	iUnitId: INT;
	//2025.10.28.140624 | bai.zy | 单运行的轴速度先单独拿出来
	adiVel_Virtual_Tar_Inch : ARRAY [1..MAX_UNIT_NUM] OF DINT;
	afbTRIG_SwitchInching_Prn: ARRAY [1..MAX_UNIT_NUM] OF R_TRIG;

	xHasAxisOnInchRunningSts : BOOL;

	diVel_Virtual_Tar_Inch_Pre : DINT;
	xHasAxisOnInchRunningSts_Pre : BOOL;

	xPrintInching_Pre : BOOL;
	xPrintInching_Lasting : BOOL;
	xInchDecing : BOOL;
	iInchDecCnt : INT;

	iDecCnt : INT;
	//2026.04.01.170415 Hou.N 增加总匀墨处理逻辑
	afbTRIG_SwitchInching_Net_On:ARRAY [1..MAX_UNIT_NUM] OF  R_TRIG;
	afbTRIG_SwitchInching_Net_Off: ARRAY [1..MAX_UNIT_NUM] OF R_TRIG;
	xSwitch_Inching_Net:ARRAY [1..MAX_UNIT_NUM] OF BOOL;
	aitest1:ARRAY [1..MAX_UNIT_NUM] OF INT;
	aitest2:ARRAY [1..MAX_UNIT_NUM] OF INT;

	fbTRIG_SwitchInching_Net_On : R_TRIG;
	fbTRIG_SwitchInching_Net_Off : R_TRIG;
	axSwitch_Inch_Net: ARRAY [1..MAX_UNIT_NUM] OF BOOL;
	aiTest:ARRAY [1..MAX_UNIT_NUM] OF INT;
	afbTRIG_Switch:ARRAY [1..MAX_UNIT_NUM] OF R_TRIG;
END_VAR

{IMPLEMENTATION}
o_lrMax_a_S_pos_Inch:= 1;
IF i_xEn THEN
	IF (i_iGrpId=1 OR i_iGrpId=2) AND
		(i_iGrpAxisNum_Pu>=1 AND i_iGrpAxisNum_Pu<=MAX_STATION_NUM) AND
		i_pstStSysParam<>0 THEN

		//2026.04.01.170603 Hou.N 增加总匀墨处理
(*		fbTRIG_SwitchInching_Net_On(CLK:=i_pstStSysParam^.astStRSV_GrpParam_UnSave[i_iGrpId].xSwitch_GrpInkEn );
		IF fbTRIG_SwitchInching_Net_On.Q THEN
			FOR iN := 1 TO i_iGrpAxisNum_Pu BY 1 DO
				IF i_pstStSysParam^.astStUnitParam_Save[iN].xLinkage THEN
					i_pstStSysParam^.astStRSV_UnitParam_UnSave[iN].xSwitch_Inching_Net :=TRUE;
				END_IF
			END_FOR
		END_IF

		fbTRIG_SwitchInching_Net_Off(CLK:= NOT i_pstStSysParam^.astStRSV_GrpParam_UnSave[i_iGrpId].xSwitch_GrpInkEn );
		IF fbTRIG_SwitchInching_Net_Off.Q THEN
			FOR iN := 1 TO i_iGrpAxisNum_Pu BY 1 DO
				IF i_pstStSysParam^.astStUnitParam_Save[iN].xLinkage THEN
					i_pstStSysParam^.astStRSV_UnitParam_UnSave[iN].xSwitch_Inching_Net :=FALSE;
				END_IF
			END_FOR
		END_IF
*)
		IF NOT i_pstStSysParam^.astStRSV_GrpParam_UnSave[i_iGrpId].xSwitch_GrpInkEn THEN
			FOR iN:=1 TO i_iGrpAxisNum_Pu BY 1 DO
				iUnitId:= i_aiGrpAxisList[iN];
				axSwitch_Inch_Net[iUnitId]:= FALSE;
			END_FOR
		ELSE
			FOR iN:=1 TO i_iGrpAxisNum_Pu BY 1 DO
				iUnitId:= i_aiGrpAxisList[iN];
				axSwitch_Inch_Net[iUnitId]:= i_pstStSysParam^.astStRSV_UnitParam_UnSave[iUnitId].xSwitch_Inching_Net;
			END_FOR
		END_IF

		FOR iN:=1 TO i_iGrpAxisNum_Pu BY 1 DO
			iUnitId:= i_aiGrpAxisList[iN];

			afbTRIG_SwitchInching_Prn[iUnitId](CLK := i_pastStIOMap_Axis_FE^[iUnitId].i_xInch );
			IF afbTRIG_SwitchInching_Prn[iUnitId].Q THEN
				//2026.09.06.103922 当前凹印机现场使用时，设备类型强制写4，也并在条件里
				IF i_pstStSysParam^.stStSysParam_Save.dwEquipmentProf.3 or i_pstStSysParam^.stStSysParam_Save.dwEquipmentProf.2 THEN //凹印机只能在单动时候使用2026.5.27.103527
				//IF i_pstStSysParam^.stStSysParam_Save.dwEquipmentProf.3 THEN //凹印机只能在单动时候使用2026.5.27.103527
					IF (NOT i_pstStSysParam^.astStUnitParam_Save[iUnitId].xLinkage) THEN
						i_pstStSysParam^.astStRSV_UnitParam_UnSave[iUnitId].xSwitch_Inching_Prn := NOT i_pstStSysParam^.astStRSV_UnitParam_UnSave[iUnitId].xSwitch_Inching_Prn;
					END_IF
				ELSE//其他机型先不限制单联动吧|只针对版辊2026.5.27.103529
					i_pstStSysParam^.astStRSV_UnitParam_UnSave[iUnitId].xSwitch_Inching_Prn := NOT i_pstStSysParam^.astStRSV_UnitParam_UnSave[iUnitId].xSwitch_Inching_Prn;
				END_IF
			END_IF

			i_pstStSysParam^.astStRSV_UnitParam_UnSave[iUnitId].xInching_NetRoller:=
				axSwitch_Inch_Net[iUnitId];
				//i_pstStSysParam^.astStRSV_UnitParam_UnSave[iUnitId].xSwitch_Inching_Net;
			i_pstStSysParam^.astStRSV_UnitParam_UnSave[iUnitId].xInching_BottomRoller:=
				i_pstStSysParam^.astStRSV_UnitParam_UnSave[iUnitId].xSwitch_Inching_Bottom;
			//2026.04.06.131959  test
			afbTRIG_Switch[iUnitId](CLK := i_pstStSysParam^.astStRSV_UnitParam_UnSave[iUnitId].xSwitch_Inching_Prn) ;
			IF 	afbTRIG_Switch[iUnitId].Q THEN
				aiTest[iUnitId]:=aiTest[iUnitId]+1;
			END_IF

			i_pstStSysParam^.astStUnitParam_UnSave[iUnitId].xAxisInching :=
				i_pstStSysParam^.astStRSV_UnitParam_UnSave[iUnitId].xSwitch_Inching_Prn;

			IF i_pstStSysParam^.astStGrpParam_UnSave[i_iGrpId].xPrintInching THEN
				i_pstStSysParam^.astStRSV_UnitParam_UnSave[iUnitId].xInching_NetRoller := TRUE;
				i_pstStSysParam^.astStRSV_UnitParam_UnSave[iUnitId].xInching_BottomRoller := TRUE;
				i_pstStSysParam^.astStUnitParam_UnSave[iUnitId].xAxisInching := TRUE;
			END_IF
		END_FOR

		//增加牵引
		i_pstStSysParam^.astStRSV_GrpParam_UnSave[i_iGrpId].xInching_If_Roller := i_pstStSysParam^.astStRSV_GrpParam_UnSave[i_iGrpId].xSwitch_Inching_If;
		i_pstStSysParam^.astStRSV_GrpParam_UnSave[i_iGrpId].xInching_Of_Roller := i_pstStSysParam^.astStRSV_GrpParam_UnSave[i_iGrpId].xSwitch_Inching_Of;
		IF i_pstStSysParam^.astStGrpParam_UnSave[i_iGrpId].xPrintInching THEN
			i_pstStSysParam^.astStRSV_GrpParam_UnSave[i_iGrpId].xInching_If_Roller :=TRUE;
		    i_pstStSysParam^.astStRSV_GrpParam_UnSave[i_iGrpId].xInching_Of_Roller :=TRUE;
		END_IF

		IF NOT i_pstStSysParam^.astStGrpParam_UnSave[i_iGrpId].xFlag_Stop OR (*非停机状态下,禁止各种形式的单运行*)
			(i_pstStEvtReq^.xReqStop AND i_pstStSysParam^.astStGrpParam_UnSave[i_iGrpId].xFlag_Stop) THEN(*2021.10.15.094231 增加按下停止按钮时候清除单运行*)
			FOR iN:=1 TO i_iGrpAxisNum_Pu BY 1 DO
				iUnitId:= i_aiGrpAxisList[iN];(*轴id|*)
				i_pstStSysParam^.astStRSV_UnitParam_UnSave[iUnitId].xInching_NetRoller:=FALSE;
				i_pstStSysParam^.astStRSV_UnitParam_UnSave[iUnitId].xInching_BottomRoller:=FALSE;
 				i_pstStSysParam^.astStUnitParam_UnSave[iUnitId].xAxisInching := FALSE;

				(*2026.09.06.103518+ 非停机状态下的单运行标志清除，否则会出现开机过程中按过单运行，停机后自动单运行*)
				i_pstStSysParam^.astStRSV_UnitParam_UnSave[iUnitId].xSwitch_Inching_Prn := FALSE;
            	i_pstStSysParam^.astStRSV_UnitParam_UnSave[iUnitId].xSwitch_Inching_Net := FALSE;
           		i_pstStSysParam^.astStRSV_UnitParam_UnSave[iUnitId].xSwitch_Inching_Bottom :=FALSE;
			END_FOR
			(*非停机的时候清除全体运行标志|2019.12.6.110407*)

			//增加牵引
			i_pstStSysParam^.astStRSV_GrpParam_UnSave[i_iGrpId].xInching_If_Roller := FALSE;
			i_pstStSysParam^.astStRSV_GrpParam_UnSave[i_iGrpId].xInching_Of_Roller := FALSE;

		END_IF
(*
		FOR iN:=1 TO i_iGrpAxisNum_Pu  BY 1 DO
			iUnitId:= i_aiGrpAxisList[iN];(*轴id|*)

			IF 	i_pstStSysParam^.astStRSV_UnitParam_UnSave[iUnitId].xInching_NetRoller OR
				i_pstStSysParam^.astStRSV_UnitParam_UnSave[iUnitId].xInching_BottomRoller OR
				i_pstStSysParam^.astStUnitParam_UnSave[iUnitId].xAxisInching THEN
	// 			IF pstStUnitParam_UnSave^.iAxisPrnRunCaseId=MOTION_STEP_Nothing THEN(*这里做速度规划-让主轴先动起来*)
					adiVel_Virtual_Tar_Inch[iUnitId] := LREAL_TO_DINT(i_pstStSysParam^.astStGrpParam_Save[i_iGrpId].rVel_Inch
																	*GC_LRMOTORPPR/
																	gc_rGirth_Master/60.0/1000);
					o_lrMax_a_S_pos_Inch:= 1;

					IF NOT o_xHasAxisOnInchRunningSts THEN
						o_xHasAxisOnInchRunningSts:= TRUE;
					END_IF
				//END_IF
			ELSE
				o_xHasAxisOnInchRunningSts:= FALSE;
				//o_diVel_Virtual_Tar_Inch:= 0;
				adiVel_Virtual_Tar_Inch[iUnitId] := 0;
				o_lrMax_a_S_pos_Inch:= 1;

			END_IF
		END_FOR

		IF i_pstStSysParam^.astStRSV_GrpParam_UnSave[i_iGrpId].xInching_If_Roller OR
			i_pstStSysParam^.astStRSV_GrpParam_UnSave[i_iGrpId].xInching_Of_Roller THEN

			adiVel_Virtual_Tar_Inch[i_iGrpId] := LREAL_TO_DINT(i_pstStSysParam^.astStGrpParam_Save[i_iGrpId].rVel_Inch
																	*GC_LRMOTORPPR/
																	gc_rGirth_Master/60.0/1000);
			o_lrMax_a_S_pos_Inch:= 1;

			//点动速度为5米/分
			IF i_pstStSysParam^.astStGrpParam_UnSave[i_iGrpId].xPrintInching THEN
				adiVel_Virtual_Tar_Inch[i_iGrpId] := LREAL_TO_DINT(i_pstStSysParam^.astStGrpParam_UnSave[i_iGrpId].rVel_Inching_Print
																	*GC_LRMOTORPPR/
																	gc_rGirth_Master/60.0/1000);
			END_IF
		END_IF
*)
		xHasAxisOnInchRunningSts := FALSE;
		FOR iN:=1 TO i_iGrpAxisNum_Pu  BY 1 DO
			iUnitId:= i_aiGrpAxisList[iN];(*轴id|*)
			IF 	i_pstStSysParam^.astStRSV_UnitParam_UnSave[iUnitId].xInching_NetRoller OR
				i_pstStSysParam^.astStRSV_UnitParam_UnSave[iUnitId].xInching_BottomRoller OR
				i_pstStSysParam^.astStUnitParam_UnSave[iUnitId].xAxisInching THEN
				xHasAxisOnInchRunningSts := TRUE;
				EXIT;
			END_IF
		END_FOR

		xHasAxisOnInchRunningSts := xHasAxisOnInchRunningSts OR
			i_pstStSysParam^.astStRSV_GrpParam_UnSave[i_iGrpId].xInching_If_Roller OR
			i_pstStSysParam^.astStRSV_GrpParam_UnSave[i_iGrpId].xInching_Of_Roller;

		IF xHasAxisOnInchRunningSts THEN
			o_diVel_Virtual_Tar_Inch := LREAL_TO_DINT(i_pstStSysParam^.astStGrpParam_Save[i_iGrpId].rVel_Inch
																	*GC_LRMOTORPPR/
																	gc_rGirth_Master/60.0/1000);
			o_lrMax_a_S_pos_Inch:= 1;
			//点动速度为5米/分
			IF i_pstStSysParam^.astStGrpParam_UnSave[i_iGrpId].xPrintInching THEN
				o_diVel_Virtual_Tar_Inch := LREAL_TO_DINT(i_pstStSysParam^.astStGrpParam_UnSave[i_iGrpId].rVel_Inching_Print
																	*GC_LRMOTORPPR/
																	gc_rGirth_Master/60.0/1000);
			END_IF
		ELSIF xHasAxisOnInchRunningSts_Pre <> xHasAxisOnInchRunningSts AND NOT xInchDecing THEN
			xInchDecing := TRUE;
			iDecCnt := REAL_TO_INT(i_pstStSysParam^.astStGrpParam_UnSave[i_iGrpId].rVel_Cur*1000/(i_rAcc_Inch*1000/gc_TENSION_TSK_CYCLE_TIME)/gc_TENSION_TSK_CYCLE_TIME+0.5);
			o_diVel_Virtual_Tar_Inch := LREAL_TO_DINT(i_pstStSysParam^.astStGrpParam_Save[i_iGrpId].rVel_Inch
																	*GC_LRMOTORPPR/
																	gc_rGirth_Master/60.0/1000);
			o_lrMax_a_S_pos_Inch:= 1;
			//点动速度为5米/分
			IF i_pstStSysParam^.astStGrpParam_UnSave[i_iGrpId].xPrintInching THEN
				o_diVel_Virtual_Tar_Inch := LREAL_TO_DINT(i_pstStSysParam^.astStGrpParam_UnSave[i_iGrpId].rVel_Inching_Print
																	*GC_LRMOTORPPR/
																	gc_rGirth_Master/60.0/1000);
			END_IF

			IF xPrintInching_Pre <>i_pstStSysParam^.astStGrpParam_UnSave[i_iGrpId].xPrintInching THEN
				xPrintInching_Lasting := TRUE;
			END_IF
		ELSIF xInchDecing THEN
			o_diVel_Virtual_Tar_Inch := LREAL_TO_DINT(i_pstStSysParam^.astStGrpParam_Save[i_iGrpId].rVel_Inch
																	*GC_LRMOTORPPR/
																	gc_rGirth_Master/60.0/1000);
			o_lrMax_a_S_pos_Inch:= 1;
			//点动速度为5米/分
			IF i_pstStSysParam^.astStGrpParam_UnSave[i_iGrpId].xPrintInching OR xPrintInching_Lasting THEN
				o_diVel_Virtual_Tar_Inch := LREAL_TO_DINT(i_pstStSysParam^.astStGrpParam_UnSave[i_iGrpId].rVel_Inching_Print
																	*GC_LRMOTORPPR/
																	gc_rGirth_Master/60.0/1000);
			END_IF
			iInchDecCnt := iInchDecCnt + 1;
			IF iInchDecCnt > iDecCnt THEN//8*1000/gc_TENSION_TSK_CYCLE_TIME THEN
				iInchDecCnt := 0;
				xInchDecing := FALSE;
				xPrintInching_Lasting := FALSE;
			END_IF
		ELSE
			o_xHasAxisOnInchRunningSts:= FALSE;	;
			//adiVel_Virtual_Tar_Inch[iUnitId] := 0;
			o_diVel_Virtual_Tar_Inch := 0;
			o_lrMax_a_S_pos_Inch:= 1;

			xInchDecing := FALSE;
			xPrintInching_Lasting := FALSE;
		END_IF
		diVel_Virtual_Tar_Inch_Pre := o_diVel_Virtual_Tar_Inch;
		xHasAxisOnInchRunningSts_Pre := xHasAxisOnInchRunningSts;
		xPrintInching_Pre := i_pstStSysParam^.astStGrpParam_UnSave[i_iGrpId].xPrintInching;
		o_xInchDecing := xInchDecing;
		//2025.10.28.140948 | bai.zy | 输出速度
// 		FOR iN := 1 TO i_iGrpAxisNum_Pu BY 1 DO
// 			iUnitId:= i_aiGrpAxisList[iN];(*轴id|*)
// 			IF (i_pstStSysParam^.astStRSV_GrpParam_UnSave[i_iGrpId].xInching_If_Roller OR i_pstStSysParam^.astStRSV_GrpParam_UnSave[i_iGrpId].xInching_Of_Roller OR
// 				i_pstStSysParam^.astStRSV_UnitParam_UnSave[iUnitId].xInching_NetRoller  OR i_pstStSysParam^.astStRSV_UnitParam_UnSave[iUnitId].xInching_BottomRoller OR i_pstStSysParam^.astStUnitParam_UnSave[iUnitId].xAxisInching) AND
// 				 adiVel_Virtual_Tar_Inch[iN] <> 0 THEN
// 				o_diVel_Virtual_Tar_Inch :=  adiVel_Virtual_Tar_Inch[iN];
// 				EXIT;
// 			END_IF
// 		END_FOR
	ELSE;
	END_IF
END_IF

(* ---- KS_FB_AxisModeCtl.st ---- *)
(*@CES
Name=KS_FB_AxisModeCtl
Type=FunctionBlock
TypeGuid=6f9dac99-8de1-4efc-8465-68ac443b7d08
Guid=88b2c618-b0a1-49ee-8cb5-d949cd68b5c9
HasDeclaration=True
HasImplementation=True
*)
{DECLARATION}
FUNCTION_BLOCK KS_FB_AxisModeCtl
VAR_INPUT
	i_xEn: BOOL;
	i_iGrpId: INT;
	i_iGrpUnitNum_Pu : INT;
	i_aiGrpUnitList: ARRAY [1..MAX_UNIT_NUM] OF INT;
	i_iGrpGearMotion_Num: INT;
	i_aiGrpGearMotion_StdList: ARRAY [1..MAX_STATION_NUM] OF INT;
	i_pstStSysParam: POINTER TO StSysParam;
	i_pastStAxisIdListInf :POINTER TO ARRAY [1..128] OF StAxisIdListInf;
	i_pastStMotorParam_Vel: POINTER TO ARRAY [1..MAX_STATION_NUM] OF StMotorParam_Vel;
	i_pstStSysStationInf			:POINTER TO StSysStationInf;
END_VAR
VAR_OUTPUT
END_VAR
VAR
	iN: INT;
	iAxisId: INT;
	iTypeId: INT;
	iUnitId: INT;
	iCoreId: INT;
	iGroupId : INT;
	iAdjAxisId : INT;
	pstStGrpParam_Save: POINTER TO StGrpParam_Save;
	pstStGrpParam_UnSave: POINTER TO StGrpParam_UnSave;

END_VAR

{IMPLEMENTATION}
IF i_xEn THEN
	IF (i_iGrpId=1 OR i_iGrpId=2) AND
		i_iGrpUnitNum_Pu>=1 AND i_iGrpUnitNum_Pu<=MAX_UNIT_NUM AND
		i_iGrpGearMotion_Num>=1 AND i_iGrpGearMotion_Num<= MAX_STATION_NUM AND
		i_pstStSysParam<>0 AND
		i_pastStAxisIdListInf<>0 AND
		i_pastStMotorParam_Vel<>0 AND
		i_pstStSysStationInf <> 0 THEN
		pstStGrpParam_Save:= ADR(i_pstStSysParam^.astStGrpParam_Save[i_iGrpId]);
		pstStGrpParam_UnSave:= ADR(i_pstStSysParam^.astStGrpParam_UnSave[i_iGrpId]);

		FOR iN:=1 TO i_iGrpGearMotion_Num BY 1 DO
// 			KS_HY_GetAxisIdForMotByStation(
// 				i_aiGrpGearMotion_StdList[iN],
// 				ADR(iAxisId),
// 				ADR(iTypeId),
// 				ADR(iUnitId),
// 				ADR(iCoreId),
// 				ADR(iGroupId),
// 				ADR(iAdjAxisId),
// 				i_pastStAxisIdListInf);
			KS_GetAxisIdForMotByStation_V2(
					i_iStationId:= i_aiGrpGearMotion_StdList[iN],
					i_piAxisId:= ADR(iAxisId),
					i_piTypeId:= ADR(iTypeId),
					i_piUnitId:= ADR(iUnitId),
					i_piCoreId:= ADR(iCoreId),
					i_piGroupId:= ADR(iGroupId),
					i_piAdjAxisId:= ADR(iAdjAxisId),
					i_pstStSysStationInf:= i_pstStSysStationInf);
			CASE iTypeId OF
			TYPE_MASTER_I,TYPE_MASTER_II:
				i_pastStMotorParam_Vel^[iN].iMotionMode:= 1;(*虚拟主轴JOG*)
			TYPE_CENTRAL_I,TYPE_CENTRAL_II:
				i_pastStMotorParam_Vel^[iN].iMotionMode:= 0;(*电子齿轮*)
			TYPE_UNWIND_A_I,TYPE_UNWIND_A_II,
			TYPE_UNWIND_B_I,TYPE_UNWIND_B_II,
			TYPE_REWIND_A_I,TYPE_REWIND_A_II,
			TYPE_REWIND_B_I,TYPE_REWIND_B_II:
				i_pastStMotorParam_Vel^[iN].iMotionMode:= 3;(*jog*)
(*2026.4.27.215845|收放料改用速度模式
			TYPE_UNWIND_A_I,TYPE_UNWIND_A_II:
				i_pastStMotorParam_Vel^[iN].iMotionMode:= 0;(*电子齿轮*)
				IF pstStGrpParam_UnSave^.xInching_Uw THEN
					i_pastStMotorParam_Vel^[iN].iMotionMode:= 1;(*收放料单运行就先按JOG走吧*)
				END_IF
			TYPE_UNWIND_B_I,TYPE_UNWIND_B_II:
				i_pastStMotorParam_Vel^[iN].iMotionMode:= 0;(*电子齿轮*)
				IF pstStGrpParam_UnSave^.xInching_Uw THEN
					i_pastStMotorParam_Vel^[iN].iMotionMode:= 1;(*收放料单运行就先按JOG走吧*)
				END_IF
			TYPE_REWIND_A_I,TYPE_REWIND_A_II:
				i_pastStMotorParam_Vel^[iN].iMotionMode:= 0;(*电子齿轮*)
				IF pstStGrpParam_UnSave^.xInching_Rw THEN
					i_pastStMotorParam_Vel^[iN].iMotionMode:= 1;(*收放料单运行就先按JOG走吧*)
				END_IF
			TYPE_REWIND_B_I,TYPE_REWIND_B_II:
				i_pastStMotorParam_Vel^[iN].iMotionMode:= 0;(*电子齿轮*)
				IF pstStGrpParam_UnSave^.xInching_Rw THEN
					i_pastStMotorParam_Vel^[iN].iMotionMode:= 1;(*收放料单运行就先按JOG走吧*)
				END_IF
*)
			TYPE_INFEED_I,TYPE_INFEED_II:
				i_pastStMotorParam_Vel^[iN].iMotionMode:= 0;(*电子齿轮*)
				IF pstStGrpParam_UnSave^.xInching_If THEN
					i_pastStMotorParam_Vel^[iN].iMotionMode:= 1;(*单运行就先按JOG走吧*)
				END_IF
			TYPE_OUTFEED_I,TYPE_OUTFEED_II:
				i_pastStMotorParam_Vel^[iN].iMotionMode:= 0;(*电子齿轮*)
				IF pstStGrpParam_UnSave^.xInching_Of THEN
					i_pastStMotorParam_Vel^[iN].iMotionMode:= 1;(*单运行就先按JOG走吧*)
				END_IF
			TYPE_UNIT_PRN:
				i_pastStMotorParam_Vel^[iN].iMotionMode:= 0;(*电子齿轮*)

				IF pstStGrpParam_UnSave^.xFlag_Home OR pstStGrpParam_UnSave^.xFlag_PreRegister OR pstStGrpParam_UnSave^.xFlag_PhaseRead OR pstStGrpParam_UnSave^.xFlag_PhaseRestore THEN
					i_pastStMotorParam_Vel^[iN].iMotionMode:= 2;(*回原点等用点位*)
				END_IF
				(*版辊单运行还是按照电子齿轮走|方便执行印刷切换单联动标志*)
				//2025.10.28.104901 | bai.zy | 增加单运行
				IF pstStGrpParam_UnSave^.xFlag_AllInchRun OR i_pstStSysParam^.astStUnitParam_UnSave[iUnitId].xAxisInching THEN
					i_pastStMotorParam_Vel^[iN].iMotionMode:= 1;(*电子齿轮*)
				END_IF

			TYPE_UNIT_BOTTOM:
				i_pastStMotorParam_Vel^[iN].iMotionMode:= 0;(*电子齿轮*)

				//柔印单伺服底辊
				IF g_iMachineryType	= MACHINERYTYPE_FELXO_INLINE_ONEBOTOMROLLER THEN
					IF pstStGrpParam_UnSave^.xFlag_Home OR pstStGrpParam_UnSave^.xFlag_PreRegister OR pstStGrpParam_UnSave^.xFlag_PhaseRead OR pstStGrpParam_UnSave^.xFlag_PhaseRestore THEN
						i_pastStMotorParam_Vel^[iN].iMotionMode:= 2;(*回原点等用点位*)
					END_IF
					(*版辊单运行还是按照电子齿轮走|方便执行印刷切换单联动标志*)
					//2025.10.28.104901 | bai.zy | 增加单运行
					IF pstStGrpParam_UnSave^.xFlag_AllInchRun OR i_pstStSysParam^.astStUnitParam_UnSave[iUnitId].xAxisInching THEN
						i_pastStMotorParam_Vel^[iN].iMotionMode:= 1;(*电子齿轮*)
					END_IF
				END_IF
			TYPE_UNIT_NET:
				i_pastStMotorParam_Vel^[iN].iMotionMode:= 0;(*电子齿轮*)
				IF i_pstStSysParam^.astStRSV_UnitParam_UnSave[iUnitId].xInching_NetRoller THEN
					i_pastStMotorParam_Vel^[iN].iMotionMode:= 1;(*电子齿轮*)
				END_IF
			END_CASE
		END_FOR
	END_IF
ELSE
	;
END_IF

(* ---- KS_FB_AxisTrapPosCtl.st ---- *)
(*@CES
Name=KS_FB_AxisTrapPosCtl
Type=FunctionBlock
TypeGuid=6f9dac99-8de1-4efc-8465-68ac443b7d08
Guid=2e2173c6-f3c4-47fe-9b59-d4fa6be54b09
HasDeclaration=True
HasImplementation=True
*)
{DECLARATION}
FUNCTION_BLOCK KS_FB_AxisTrapPosCtl(*预套准、相位回复等位置计0算*)
VAR_INPUT
	i_xEn: BOOL;
	i_iGrpId: INT;
	i_iGrpAxisNum_Pu: INT;
	i_aiGrpUnitList: ARRAY [1..MAX_UNIT_NUM] OF INT;
	i_pstStSysParam: POINTER TO StSysParam;
//	i_pastStWatch_Sts_display_Prn				: POINTER TO ARRAY [1..MAX_UNIT_NUM] OF StWatch_Sts_display;
	//i_pastStWatch_Sts_display_Bottom			: POINTER TO ARRAY [1..MAX_UNIT_NUM] OF StWatch_Sts_display;
	i_pawAxisVirtualCnt: POINTER TO ARRAY [1..MAX_UNIT_NUM] OF WORD; (* 2021.6.25.104504/增加的虚拟编码器原始值输入 *)
	i_pawAxisVirtualSts: POINTER TO ARRAY [1..MAX_UNIT_NUM] OF WORD; (* 2021.6.25.104504/增加的虚拟编码器原始值输入 *)
	i_diTime_PreReg: DINT:=5000;//5s内走完

	i_padiPreRegisterPos: POINTER TO ARRAY [1..MAX_UNIT_NUM] OF DINT;
	i_palrMaxVel_PreReg: POINTER TO ARRAY [1..MAX_UNIT_NUM] OF LREAL;//预套准最大速度-时间固定，速度不同
	//2024.10.22.193803增加单圈绝对位置计算预套准
	//i_padiEncPos_Virtual_start_0: POINTER TO ARRAY [1..MAX_UNIT_NUM] OF DINT;
	i_pastStGetMotionSts: POINTER TO ARRAY [1..MAX_STATION_NUM] OF StGetMotionSts;
	i_pstStSysStationInf			:POINTER TO StSysStationInf;
END_VAR
VAR_OUTPUT
	o_xEn: BOOL;
END_VAR
VAR
	fbRTrig_Home: R_TRIG;
	fbRTrig_PreRegister: R_TRIG;
	fbRTrig_PhaseRestore: R_TRIG;
	xCalcAdjustPos: BOOL:= FALSE;
	iN: INT;
	iUnitId:INT;
	pstStGrpParam_Save: POINTER TO StGrpParam_Save;
	pstStGrpParam_UnSave: POINTER TO StGrpParam_UnSave;
	pstStUnitParam_Save: POINTER TO StUnitParam_Save;
	pstStUnitParam_UnSave: POINTER TO StUnitParam_UnSave;
	lrMotorPPR_temp: LREAL;
	alrMotorNeedMovePos_Pul: ARRAY [1..MAX_UNIT_NUM] OF LREAL;
	alrAxisMotorPulseMovement: ARRAY [1..MAX_UNIT_NUM] OF LREAL;

	xFlag_PreRegValueReloaded: BOOL;
	axVirEncOffsetInitialized: ARRAY [1..MAX_UNIT_NUM] OF BOOL;
	iTemp: INT;
	alrMaxVel_PreReg: ARRAY [1..MAX_UNIT_NUM] OF LREAL;//预套准最大速度-时间固定，速度不同
	alrMotorNeedMovePos_Temp_PreReg_test: ARRAY [1..MAX_UNIT_NUM] OF LREAL;
	iDeltaPhase_MarkPos_FirstLinkage: INT;
	iTmp: INT;
	wVirtuaCnt_Temp: WORD;

	iAxisId : INT;
	xFlag_PreReg:BOOL;
	xFlag_PreReg_End:BOOL;
	iTimeCnt: INT;

	lrTmp : LREAL;
	lrTmp1 : LREAL;
	rMaxAdjust : REAL;
	rAcc_TargetAxis : REAL := 2.0;
	rTime_Acc : REAL;
	arTargetVel : ARRAY [1..MAX_UNIT_NUM] OF REAL;
	xFlag_PreReg_Finished : BOOL;

	iTypeId: INT;
	iCoreId: INT;
	iGroupId : INT;
	iAdjAxisId : INT;
END_VAR

{IMPLEMENTATION}
IF i_xEn THEN
	IF	i_pstStSysParam<>0 AND i_iGrpAxisNum_Pu>=1 AND i_iGrpAxisNum_Pu<=MAX_UNIT_NUM  AND
		 i_pawAxisVirtualCnt<>0 AND i_padiPreRegisterPos<>0 AND i_palrMaxVel_PreReg<>0AND
		i_diTime_PreReg<>0 AND i_pastStGetMotionSts <> 0 THEN
		pstStGrpParam_Save:= ADR(i_pstStSysParam^.astStGrpParam_Save[i_iGrpId]);
		pstStGrpParam_UnSave:= ADR(i_pstStSysParam^.astStGrpParam_UnSave[i_iGrpId]);
		fbRTrig_Home(CLK:= pstStGrpParam_UnSave^.xFlag_Home);
		fbRTrig_PreRegister(CLK:= pstStGrpParam_UnSave^.xFlag_PreRegister);
		fbRTrig_PhaseRestore(CLK:= pstStGrpParam_UnSave^.xFlag_PhaseRestore);

		IF fbRTrig_Home.Q OR fbRTrig_PreRegister.Q OR fbRTrig_PhaseRestore.Q THEN
			IF pstStGrpParam_UnSave^.xFlag_Home THEN
				pstStGrpParam_UnSave^.xFlag_Home_end:= FALSE;
			ELSIF pstStGrpParam_UnSave^.xFlag_PreRegister THEN
				pstStGrpParam_UnSave^.xFlag_PreRegister_end:= FALSE;
			ELSIF pstStGrpParam_UnSave^.xFlag_PhaseRestore THEN
				pstStGrpParam_UnSave^.xFlag_PhaseRestore_end:= FALSE;
			END_IF

			xCalcAdjustPos:= TRUE;
		END_IF

		IF (NOT pstStGrpParam_UnSave^.xFlag_Home) AND
			(NOT pstStGrpParam_UnSave^.xFlag_PreRegister) AND
			(NOT pstStGrpParam_UnSave^.xFlag_PhaseRestore) THEN
			xFlag_PreRegValueReloaded:= FALSE;
			FOR iN:=1 TO i_iGrpAxisNum_Pu BY 1 DO
				iUnitId:= i_aiGrpUnitList[iUnitId];
				axVirEncOffsetInitialized[iUnitId]:=FALSE;
			END_FOR
		END_IF

		IF xCalcAdjustPos THEN
			xCalcAdjustPos:= FALSE;//只计算一次2023.08.11.180238
			FOR iN:=1 TO i_iGrpAxisNum_Pu BY 1 DO
				iUnitId:= i_aiGrpUnitList[iN];
				pstStUnitParam_Save:= ADR(i_pstStSysParam^.astStUnitParam_Save[iUnitId]);
				pstStUnitParam_UnSave:= ADR(i_pstStSysParam^.astStUnitParam_UnSave[iUnitId]);
				IF pstStGrpParam_UnSave^.xFlag_Home THEN
					IF pstStUnitParam_Save^.xLinkage THEN(*只计算联动轴|2022.9.8.120509*)
						//2026.1.6.134228 | + | 不同机器类型处理
						IF g_iMachineryType	= MACHINERYTYPE_FELXO_INLINE_ONEBOTOMROLLER THEN
							IF pstStUnitParam_UnSave^.xMotRev_BottomRoller THEN
								lrMotorPPR_temp:= -(GC_LRMOTORPPR)* pstStUnitParam_Save^.rGirth_PrnRoller *pstStUnitParam_Save^.uiNum_BottomRoller / pstStUnitParam_Save^.uiDen_BottomRoller/pstStUnitParam_Save^.rGirth_BottomRoller;
							ELSE
								lrMotorPPR_temp:= (GC_LRMOTORPPR)* pstStUnitParam_Save^.rGirth_PrnRoller *pstStUnitParam_Save^.uiNum_BottomRoller / pstStUnitParam_Save^.uiDen_BottomRoller/pstStUnitParam_Save^.rGirth_BottomRoller;
							END_IF
						ELSE
							IF pstStUnitParam_UnSave^.xMotRev_PrnRoller THEN
								lrMotorPPR_temp:= -(GC_LRMOTORPPR)* pstStUnitParam_Save^.uiNum_PrnRoller / pstStUnitParam_Save^.uiDen_PrnRoller;
							ELSE
								lrMotorPPR_temp:= (GC_LRMOTORPPR)* pstStUnitParam_Save^.uiNum_PrnRoller / pstStUnitParam_Save^.uiDen_PrnRoller;
							END_IF
						END_IF

						alrMotorNeedMovePos_Pul[iUnitId]:=lrMotorPPR_temp;
						alrMotorNeedMovePos_Pul[iUnitId]:=lrMotorPPR_temp*2;
					END_IF
				(*2017-09-13 13:26:39|
				/.预套准
				*)
				ELSIF pstStGrpParam_UnSave^.xFlag_PreRegister THEN
					IF NOT xFlag_PreRegValueReloaded THEN
						KS_ReloadPreRegValue(
							i_iGrpId,
							i_iGrpAxisNum_Pu,
							i_aiGrpUnitList,
							i_pstStSysParam,
							i_pawAxisVirtualCnt,
							i_pawAxisVirtualSts,
							ADR(alrAxisMotorPulseMovement),
							ADR(iDeltaPhase_MarkPos_FirstLinkage));
						xFlag_PreRegValueReloaded:= TRUE;
					END_IF

					IF pstStGrpParam_Save^.xPreRegisterAxisId_Manu THEN(*预套准id手动选择@2025.1.12.193735*)
						IF pstStUnitParam_Save^.xPreRegisterValid_Manu AND(*有效了@则进行预套*)
							pstStUnitParam_Save^.xLinkage THEN
							alrMotorNeedMovePos_Pul[iUnitId]:=alrAxisMotorPulseMovement[iUnitId];
						END_IF
					ELSE
						IF pstStUnitParam_Save^.xLinkage THEN(*只计算联动轴|2022.9.8.120509*)
							alrMotorNeedMovePos_Pul[iUnitId]:=alrAxisMotorPulseMovement[iUnitId];
						END_IF
					END_IF

				(*2017-09-13 13:26:58|
				/.相位恢复
				*)
				ELSIF pstStGrpParam_UnSave^.xFlag_PhaseRestore THEN
					IF pstStUnitParam_Save^.xLinkage THEN(*只计算联动轴|2022.9.8.120509*)
						//IF NOT axVirEncOffsetInitialized[iUnitId] THEN
(*deprecated@2021.6.25.113401
							IF i_pastStPTSts^[iAxisId].virtualCnt>= pstStAxisParam^.iPhase_RegisterOk THEN (*当前位置在相位点之后|那么移动的是一个补值*)
								iTemp:= (pstStAxisParam^.iPhase_RegisterOk-i_pastStPTSts^[iAxisId].virtualCnt+gc_iVirEncPPR);
with/
*)
							IF i_pawAxisVirtualCnt^[iUnitId] >= pstStUnitParam_Save^.iPhase_RegisterOk THEN (* 2021.6.25.113420/ *)
								iTemp:= (pstStUnitParam_Save^.iPhase_RegisterOk - i_pawAxisVirtualCnt^[iUnitId] + gc_iVirEncPPR); (* 2021.6.25.113649/ *)
								WHILE iTemp<0 DO
									iTemp:= iTemp+gc_iVirEncPPR;
								END_WHILE
								//2026.1.6.134228 | + | 不同机器类型处理
								IF g_iMachineryType	= MACHINERYTYPE_FELXO_INLINE_ONEBOTOMROLLER THEN
									alrAxisMotorPulseMovement[iUnitId]:= (INT_TO_LREAL(iTemp) / gc_iVirEncPPR) * ((GC_LRMOTORPPR) * pstStUnitParam_Save^.rGirth_PrnRoller *pstStUnitParam_Save^.uiNum_BottomRoller / pstStUnitParam_Save^.uiDen_BottomRoller/pstStUnitParam_Save^.rGirth_BottomRoller );
								ELSE
									alrAxisMotorPulseMovement[iUnitId]:= (INT_TO_LREAL(iTemp) / gc_iVirEncPPR) * ((GC_LRMOTORPPR) * pstStUnitParam_Save^.uiNum_PrnRoller / pstStUnitParam_Save^.uiDen_PrnRoller);
								END_IF
							ELSE (*还没到相位点*)
(*deprecated@2021.6.25.113607
								iTemp:= pstStAxisParam^.iPhase_RegisterOk-i_pastStPTSts^[iAxisId].virtualCnt;
with/
*)
								iTemp:= pstStUnitParam_Save^.iPhase_RegisterOk-i_pawAxisVirtualCnt^[iUnitId]; (* 2021.6.25.113644/ *)
								WHILE iTemp>gc_iVirEncPPR DO
									iTemp:= iTemp-gc_iVirEncPPR;
								END_WHILE
								//2026.1.6.135139 | + | 不同机器类型处理
								IF g_iMachineryType	= MACHINERYTYPE_FELXO_INLINE_ONEBOTOMROLLER THEN
									alrAxisMotorPulseMovement[iUnitId]:= (INT_TO_LREAL(iTemp) / gc_iVirEncPPR) * ((GC_LRMOTORPPR) * pstStUnitParam_Save^.rGirth_PrnRoller *pstStUnitParam_Save^.uiNum_BottomRoller / pstStUnitParam_Save^.uiDen_BottomRoller/pstStUnitParam_Save^.rGirth_BottomRoller );
								ELSE
									alrAxisMotorPulseMovement[iUnitId]:= (INT_TO_LREAL(iTemp) / gc_iVirEncPPR) * ((GC_LRMOTORPPR) * pstStUnitParam_Save^.uiNum_PrnRoller / pstStUnitParam_Save^.uiDen_PrnRoller);
								END_IF
							END_IF
							//2026.1.6.135139 | + | 不同机器类型处理
							IF g_iMachineryType	= MACHINERYTYPE_FELXO_INLINE_ONEBOTOMROLLER THEN
								IF pstStUnitParam_UnSave^.xMotRev_BottomRoller THEN
									alrAxisMotorPulseMovement[iUnitId]:= -alrAxisMotorPulseMovement[iUnitId];
								ELSE;
								END_IF
							ELSE
								IF pstStUnitParam_UnSave^.xMotRev_PrnRoller THEN
									alrAxisMotorPulseMovement[iUnitId]:= -alrAxisMotorPulseMovement[iUnitId];
								ELSE;
								END_IF
							END_IF
							axVirEncOffsetInitialized[iUnitId]:= TRUE;
						END_IF
						alrMotorNeedMovePos_Pul[iUnitId]:=alrAxisMotorPulseMovement[iUnitId];
					//END_IF
(*
				ELSIF i_pxFlag_CphCommonVir^ THEN(*通用相位初始装版相位记录*)
					FOR iN:=1 TO i_iGrpAxisNum_Pu BY 1 DO
						iAxisId:= i_aiGrpAxisList[iN];
						//pstStAxisParam:= ADR(i_pstStShmGlobalParam^.astStAxisParam[iAxisId]);
						IF i_pstStSysParam^.astStUnitParam_Save[iAxisId].xServoOn AND
							i_pstStSysParam^.astStUnitParam_Save[iAxisId].xLinkage THEN(*只计算联动轴|2022.9.8.120509*)
							IF i_pstStSysParam^.astStUnitParam_UnSave[iAxisId].xMotRev_PrnRoller THEN
								lrMotorPPR_temp:= -DWORD_TO_LREAL(gc_dwMotorPPR)* i_pstStSysParam^.astStUnitParam_Save[iAxisId].uiNum_PrnRoller / i_pstStSysParam^.astStUnitParam_Save[iAxisId].uiDen_PrnRoller;
							ELSE
								lrMotorPPR_temp:= DWORD_TO_LREAL(gc_dwMotorPPR)* i_pstStSysParam^.astStUnitParam_Save[iAxisId].uiNum_PrnRoller / i_pstStSysParam^.astStUnitParam_Save[iAxisId].uiDen_PrnRoller;
							END_IF
							alrMotorNeedMovePos_Pul[iAxisId]:=lrMotorPPR_temp;
						END_IF
					END_FOR
				ELSIF i_pxCphaseRestore^ THEN(*通用相位恢复*)
					FOR iN:=1 TO i_iGrpAxisNum_Pu BY 1 DO
						iAxisId:= i_aiGrpAxisList[iN];
						//pstStAxisParam:= ADR(i_pstStShmGlobalParam^.astStAxisParam[iAxisId]);
						IF i_pstStSysParam^.astStUnitParam_Save[iAxisId].xServoOn AND
							i_pstStSysParam^.astStUnitParam_Save[iAxisId].xLinkage THEN(*只计算联动轴|2022.9.8.120509*)
							IF NOT axVirEncOffsetInitialized[iAxisId] THEN
								iTemp:= i_pstStSysParam^.astStUnitParam_Save[iAxisId].iPhase_FinalUsed;
								alrAxisMotorPulseMovement[iAxisId]:= (INT_TO_LREAL(iTemp) / gc_iVirEncPPR) * (DWORD_TO_LREAL(gc_dwMotorPPR) * pstStAxisParam^.uiNum / pstStAxisParam^.uiDen);
								axVirEncOffsetInitialized[iAxisId]:= TRUE;
								IF i_pstStSysParam^.astStUnitParam_UnSave[iAxisId].xMotRev_PrnRoller THEN
									alrAxisMotorPulseMovement[iAxisId]:= -alrAxisMotorPulseMovement[iAxisId];
								ELSE;
								END_IF
							END_IF
							alrMotorNeedMovePos_Pul[iAxisId]:=alrAxisMotorPulseMovement[iAxisId];
						END_IF
					END_FOR
					*)
				ELSIF pstStGrpParam_Save^.xFlag_PhaseRead THEN(*固定相位恢复|2024.9.6.214324*)
					IF pstStUnitParam_Save^.xLinkage THEN(*只计算联动轴|2022.9.8.120509*)
						IF NOT axVirEncOffsetInitialized[iUnitId] THEN
							iTmp:=KS_GetPhaseValue(i_pawAxisVirtualCnt^[iUnitId],gc_iVirEncPPR);(*2023.6.28.113035 更新*)
							wVirtuaCnt_Temp:=INT_TO_WORD(iTmp);
							IF wVirtuaCnt_Temp >= pstStUnitParam_Save^.iPhase_Locating THEN (* 2021.6.25.113420/ *)
								iTemp:= (pstStUnitParam_Save^.iPhase_Locating - wVirtuaCnt_Temp + gc_iVirEncPPR); (* 2021.6.25.113649/ *)
								WHILE iTemp<0 DO
									iTemp:= iTemp+gc_iVirEncPPR;
								END_WHILE
								//2026.1.6.135139 | + | 不同机器类型处理
								IF g_iMachineryType	= MACHINERYTYPE_FELXO_INLINE_ONEBOTOMROLLER THEN
									alrAxisMotorPulseMovement[iUnitId]:= (INT_TO_LREAL(iTemp) / gc_iVirEncPPR) * ((GC_LRMOTORPPR) * pstStUnitParam_Save^.rGirth_PrnRoller * pstStUnitParam_Save^.uiNum_BottomRoller / pstStUnitParam_Save^.uiDen_BottomRoller/pstStUnitParam_Save^.rGirth_BottomRoller);
								ELSE
									alrAxisMotorPulseMovement[iUnitId]:= (INT_TO_LREAL(iTemp) / gc_iVirEncPPR) * ((GC_LRMOTORPPR) * pstStUnitParam_Save^.uiNum_PrnRoller / pstStUnitParam_Save^.uiDen_PrnRoller);
								END_IF

							ELSE (*还没到相位点*)
								iTemp:= pstStUnitParam_Save^.iPhase_Locating-wVirtuaCnt_Temp; (* 2021.6.25.113644/ *)
								WHILE iTemp>gc_iVirEncPPR DO
									iTemp:= iTemp-gc_iVirEncPPR;
								END_WHILE
								//2026.1.6.135139 | + | 不同机器类型处理
								IF g_iMachineryType	= MACHINERYTYPE_FELXO_INLINE_ONEBOTOMROLLER THEN
									alrAxisMotorPulseMovement[iUnitId]:= (INT_TO_LREAL(iTemp) / gc_iVirEncPPR) * ((GC_LRMOTORPPR) * pstStUnitParam_Save^.rGirth_PrnRoller * pstStUnitParam_Save^.uiNum_BottomRoller / pstStUnitParam_Save^.uiDen_BottomRoller/pstStUnitParam_Save^.rGirth_BottomRoller);
								ELSE
									alrAxisMotorPulseMovement[iUnitId]:= (INT_TO_LREAL(iTemp) / gc_iVirEncPPR) * ((GC_LRMOTORPPR) * pstStUnitParam_Save^.uiNum_PrnRoller / pstStUnitParam_Save^.uiDen_PrnRoller);
								END_IF

							END_IF
							//2026.1.6.135139 | + | 不同机器类型处理
							IF g_iMachineryType	= MACHINERYTYPE_FELXO_INLINE_ONEBOTOMROLLER THEN
								IF pstStUnitParam_UnSave^.xMotRev_BottomRoller THEN
									alrAxisMotorPulseMovement[iUnitId]:= -alrAxisMotorPulseMovement[iUnitId];
								ELSE;
								END_IF
							ELSE
								IF pstStUnitParam_UnSave^.xMotRev_PrnRoller THEN
									alrAxisMotorPulseMovement[iUnitId]:= -alrAxisMotorPulseMovement[iUnitId];
								ELSE;
								END_IF
							END_IF

							axVirEncOffsetInitialized[iUnitId]:= TRUE;
						END_IF
						alrMotorNeedMovePos_Pul[iUnitId]:=alrAxisMotorPulseMovement[iUnitId];
					END_IF
				ELSE;
				END_IF
(*
				(*预套时间计算*)
				(*参数单位切换*)
				IF i_pstStSysParam^.astStUnitParam_Save[iAxisId].rGirth_PrnRoller<>0 AND i_pstStSysParam^.astStUnitParam_Save[iAxisId].uiDen_PrnRoller<>0 THEN
					alrPreRegisterVel_PPMS[iAxisId]:=INT_TO_LREAL(i_iPreRegisterVel_Max)/i_pstStSysParam^.astStUnitParam_Save[iAxisId].rGirth_PrnRoller/60
													*i_pstStSysParam^.astStUnitParam_Save[iAxisId].uiNum_PrnRoller / i_pstStSysParam^.astStUnitParam_Save[iAxisId].uiDen_PrnRoller*gc_dwMotorPPR;(*电机侧速度|Pul/ms*)
				END_IF

				lrTemp:=0;
				IF alrPreRegisterVel_PPMS[iAxisId]<>0 THEN
					lrTemp:=ABS(alrMotorNeedMovePos_Pul[iAxisId])/alrPreRegisterVel_PPMS[iAxisId];(*计算最大速度匀速运动时间|MS*)
					IF lrTemp>i_iAccTime_MaxVel THEN(*超过了最大速度的加速时间|规划为梯形规划*)
						(*计算实际运动的时间*)
						(*最大速度不变*)
						lrTemp:=lrTemp+i_iAccTime_MaxVel;
						IF alrMotorNeedMovePos_Pul[iAxisId]<0 THEN(*位置小于0速度取反*)
							alrPreRegisterVel_PPMS[iAxisId]:=-alrPreRegisterVel_PPMS[iAxisId];
						END_IF
					ELSIF lrTemp>0 THEN(*规划为不能达到最大速度的三角形规划*)
						(*最大速度被改变了*)
						lrTemp:=i_iAccTime_MaxVel*2;
						IF i_iAccTime_MaxVel<>0 THEN
							alrPreRegisterVel_PPMS[iAxisId]:=(alrMotorNeedMovePos_Pul[iAxisId])/i_iAccTime_MaxVel;
						END_IF
					END_IF
				END_IF

				alrPreRegisterTime_Ms[iAxisId]:=lrTemp;
				*)
				i_padiPreRegisterPos^[iUnitId]:= LREAL_TO_DINT(alrMotorNeedMovePos_Pul[iUnitId]);
				//2025.11.13.191045 | + | 速度计算不对，应该是要计算最大速度，不是平均速度
				//i_palrMaxVel_PreReg^[iUnitId]:= ABS(alrMotorNeedMovePos_Pul[iUnitId])/i_diTime_PreReg;
				rAcc_TargetAxis := 2.0;
				rMaxAdjust:= 0.5*0.5*rAcc_TargetAxis*DINT_TO_REAL(i_diTime_PreReg)*DINT_TO_REAL(i_diTime_PreReg);
				IF ABS(alrMotorNeedMovePos_Pul[iUnitId])>rMaxAdjust THEN
					IF 	alrMotorNeedMovePos_Pul[iUnitId]>0 THEN
						alrMotorNeedMovePos_Pul[iUnitId]:= rMaxAdjust;
					ELSE
						alrMotorNeedMovePos_Pul[iUnitId]:= -rMaxAdjust;
					END_IF
					rTime_Acc:= DINT_TO_REAL(i_diTime_PreReg)*0.5;
					arTargetVel[iUnitId]:=rAcc_TargetAxis*rTime_Acc;
				ELSE
(*
					//知道调整量和调整时间，计算调整速度和加速度
					//S = a*t*t/4;
					//a = s*4/t/t;
					//v = at;
					arAcc_Out[iUnitId] := arTargetPos_Out[iUnitId]*4/arTime_Cycle[iUnitId]/arTime_Cycle[iUnitId];
					arTargetVel_Out[iUnitId] := arAcc_Out[iUnitId] * arTime_Cycle[iUnitId]*0.5 + 0.5;
*)
				(*计算最大速度*)
				(*一元二次方程x=(-b+SQRT(b²-4ac))/2a*)
				(*调整量计算公式
				arTargetPos_Out=(arTime_Cycle+arTime_Cycle-2*rTime_Acc)*rAcc_TargetAxis_In_Out*rTime_Acc*0.5*)
					lrTmp1:= ABS(alrMotorNeedMovePos_Pul[iUnitId]);
					lrTmp:= (REAL_TO_LREAL(rAcc_TargetAxis)*REAL_TO_LREAL(rAcc_TargetAxis)*
						DINT_TO_LREAL(i_diTime_PreReg*i_diTime_PreReg));
					lrTmp:= lrTmp-	REAL_TO_LREAL(4*(rAcc_TargetAxis)*lrTmp1);
					lrTmp:= SQRT(lrTmp);
					lrTmp:= -1*rAcc_TargetAxis*DINT_TO_LREAL(i_diTime_PreReg)+lrTmp;
					rTime_Acc:= lrTmp/(-2*rAcc_TargetAxis);
					arTargetVel[iUnitId]:=rAcc_TargetAxis*rTime_Acc;
				END_IF
				i_palrMaxVel_PreReg^[iUnitId]:=arTargetVel[iUnitId];

			END_FOR
		END_IF

		//2025.10.29.162354 | bai.zy |
		IF (pstStGrpParam_UnSave^.xFlag_Home OR pstStGrpParam_UnSave^.xFlag_PreRegister OR pstStGrpParam_UnSave^.xFlag_PhaseRestore) THEN
			FOR iN:=1 TO i_iGrpAxisNum_Pu BY 1 DO
				KS_GetAxisIdForMotByStation_V2(
					i_iStationId:= i_pstStSysParam^.astStUnitParam_Save[iN].iStationId,
					i_piAxisId:= ADR(iAxisId),
					i_piTypeId:= ADR(iTypeId),
					i_piUnitId:= ADR(iUnitId),
					i_piCoreId:= ADR(iCoreId),
					i_piGroupId:= ADR(iGroupId),
					i_piAdjAxisId:= ADR(iAdjAxisId),
					i_pstStSysStationInf:= i_pstStSysStationInf);
				IF NOT xFlag_PreReg THEN
					IF i_pastStGetMotionSts^[iAxisId].dwMotionSts.10 AND
						i_pastStGetMotionSts^[iAxisId].dwMotionSts.9 THEN
						xFlag_PreReg:= TRUE;//预套准/回复相位等已经开始动作
						EXIT;
					END_IF
				END_IF
			END_FOR

			IF xFlag_PreReg THEN
				xFlag_PreReg_End:= TRUE;
				FOR iN:=1 TO i_iGrpAxisNum_Pu BY 1 DO
					KS_GetAxisIdForMotByStation_V2(
						i_iStationId:= i_pstStSysParam^.astStUnitParam_Save[iN].iStationId,
						i_piAxisId:= ADR(iAxisId),
						i_piTypeId:= ADR(iTypeId),
						i_piUnitId:= ADR(iUnitId),
						i_piCoreId:= ADR(iCoreId),
						i_piGroupId:= ADR(iGroupId),
						i_piAdjAxisId:= ADR(iAdjAxisId),
						i_pstStSysStationInf:= i_pstStSysStationInf);
					IF i_pastStGetMotionSts^[iAxisId].dwMotionSts.10 AND
						i_pstStSysParam^.astStUnitParam_Save[iN].xLinkage THEN
						xFlag_PreReg_End:= FALSE;
						EXIT;
					END_IF
				END_FOR
			END_IF
			//2025.11.14.145703 | 判断运动状态然后下使能
			IF xFlag_PreReg THEN
				FOR iN:=1 TO i_iGrpAxisNum_Pu BY 1 DO
					KS_GetAxisIdForMotByStation_V2(
						i_iStationId:= i_pstStSysParam^.astStUnitParam_Save[iN].iStationId,
						i_piAxisId:= ADR(iAxisId),
						i_piTypeId:= ADR(iTypeId),
						i_piUnitId:= ADR(iUnitId),
						i_piCoreId:= ADR(iCoreId),
						i_piGroupId:= ADR(iGroupId),
						i_piAdjAxisId:= ADR(iAdjAxisId),
						i_pstStSysStationInf:= i_pstStSysStationInf);
					IF i_pastStGetMotionSts^[iAxisId].dwMotionSts.10 AND
						i_pstStSysParam^.astStUnitParam_Save[iN].xLinkage THEN
						EXIT;
					END_IF

					IF iN = i_iGrpAxisNum_Pu THEN
						xFlag_PreReg_Finished := TRUE;
					END_IF
				END_FOR
			END_IF

			iTimeCnt:= iTimeCnt+1;
			IF (xFlag_PreReg_End OR iTimeCnt>(i_diTime_PreReg+1000)/gc_TENSION_TSK_CYCLE_TIME) AND xFlag_PreReg_Finished THEN
				(*IF xFlag_PreReg_End THEN*)
				IF pstStGrpParam_UnSave^.xFlag_Home THEN
					pstStGrpParam_UnSave^.xFlag_Home:= FALSE;
					pstStGrpParam_UnSave^.xFlag_Home_end:= TRUE;
				ELSIF pstStGrpParam_UnSave^.xFlag_PreRegister THEN
					pstStGrpParam_UnSave^.xFlag_PreRegister:= FALSE;
					pstStGrpParam_UnSave^.xFlag_PreRegister_end:=TRUE;
				ELSIF pstStGrpParam_UnSave^.xFlag_PhaseRestore THEN
					pstStGrpParam_UnSave^.xFlag_PhaseRestore:= FALSE;
					pstStGrpParam_UnSave^.xFlag_PhaseRestore_end:=TRUE;
				END_IF
				(*END_IF*)

			END_IF
		ELSE
			iTimeCnt:= 0;
			xFlag_PreReg_End:= FALSE;
			xFlag_PreReg:=FALSE;
			xFlag_PreReg_Finished := FALSE;
		END_IF
	END_IF
END_IF

(* ---- KS_FB_AxisVelCtl.st ---- *)
(*@CES
Name=KS_FB_AxisVelCtl
Type=FunctionBlock
TypeGuid=6f9dac99-8de1-4efc-8465-68ac443b7d08
Guid=151c0b62-81a2-453f-8398-cdb757e1a3a2
HasDeclaration=True
HasImplementation=True
*)
{DECLARATION}
FUNCTION_BLOCK KS_FB_AxisVelCtl
VAR_INPUT
	i_xEn: BOOL;
	i_iGrpId: INT;
	i_iGrpUnitNum_Pu : INT;
	i_aiGrpUnitList: ARRAY [1..MAX_UNIT_NUM] OF INT;
	i_iGrpGearMotion_Num: INT;
	i_aiGrpGearMotion_StdList: ARRAY [1..MAX_STATION_NUM] OF INT;
	i_pstStSysParam: POINTER TO StSysParam;
	i_pastStAxisIdListInf :POINTER TO ARRAY [1..128] OF StAxisIdListInf;
	i_pastStMotorParam_Vel: POINTER TO ARRAY [1..MAX_STATION_NUM] OF StMotorParam_Vel;
	i_pastStIOMap_Main_FE						: POINTER TO ARRAY [1..4] OF StIOMap_Main_FE;(*轴io数据区域|AB系*)
	i_pastStIOMap_Axis_FE					: POINTER TO ARRAY [1..MAX_UNIT_NUM] OF StIOMap_Axis_FE;(*轴io数据区域|`````````````````````````````````````````````*)
	i_xMotionEnabled: BOOL;(*|2021.1.15.092801 速度控制块使能修改为输入输出变量|这里处理该值的复位*)
	i_pstStSysStationInf			:POINTER TO StSysStationInf;
//2026.5.9.220343
	//增加加速度及加加速度输入只2026.4.11.153755
	i_paxFlag_PressDne: POINTER TO ARRAY [1..MAX_UNIT_NUM] OF BOOL;
	i_rVel_A: REAL;//加速度
	i_rVel_Jerk: REAL;//加加速度；
END_VAR
VAR_OUTPUT
END_VAR
VAR
	iN: INT;
	iAxisId: INT;
	iTypeId: INT;
	iUnitId: INT;
	iCoreId: INT;
	iGroupId : INT;
	iAdjAxisId : INT;
	pstStGrpParam_Save: POINTER TO StGrpParam_Save;
	pstStGrpParam_UnSave: POINTER TO StGrpParam_UnSave;
	fbKS_FB_AxisVelCtl_PrnRoller: KS_FB_AxisVelCtl_PrnRoller;
	alrAxisMotionVel:ARRAY [1..MAX_UNIT_NUM] OF LREAL;(*轴的速度值*)
	lrTempAxisVel: LREAL;(**)
//2026.5.9.220120速度升速补偿
	fbKS_FB_Compensate_Vel_Prn: KS_FB_Compensate_Vel_Prn;
	aiGrpLinkageAxisList: ARRAY [1..MAX_UNIT_NUM] OF INT;
	arAxisVelPrf_Coeff1: ARRAY [1..MAX_UNIT_NUM] OF REAL;
	arAxisVelPrf_Coeff2: ARRAY [1..MAX_UNIT_NUM] OF REAL;
	arAxisVelPrf_Coeff3: ARRAY [1..MAX_UNIT_NUM] OF REAL;
	alrAxisPrfVel: ARRAY [1..MAX_UNIT_NUM] OF LREAL;
END_VAR

{IMPLEMENTATION}
IF i_xEn THEN
	IF (i_iGrpId=1 OR i_iGrpId=2) AND
		i_iGrpUnitNum_Pu>=1 AND i_iGrpUnitNum_Pu<=MAX_UNIT_NUM AND
		i_iGrpGearMotion_Num>=1 AND i_iGrpGearMotion_Num<= MAX_STATION_NUM AND
		i_pstStSysParam<>0 AND
		i_pastStAxisIdListInf<>0 AND
		i_pastStMotorParam_Vel<>0 AND
		i_pstStSysStationInf <>0 THEN
		pstStGrpParam_Save:= ADR(i_pstStSysParam^.astStGrpParam_Save[i_iGrpId]);
		pstStGrpParam_UnSave:= ADR(i_pstStSysParam^.astStGrpParam_UnSave[i_iGrpId]);

//2026.04.11.204947
		FOR iN:=1 TO g_aiGrpLinkageAxisNum_Pu[i_iGrpId] BY 1 DO
			aiGrpLinkageAxisList[iN]:= g_aiGrpLinkageAxisList[i_iGrpId,iN];
		END_FOR

		FOR iN:=1 TO  i_iGrpUnitNum_Pu BY 1 DO
			iUnitId:= i_aiGrpUnitList[iN];
			arAxisVelPrf_Coeff1[iUnitId]:= i_pstStSysParam^.astStUnitParam_Save[iUnitId].rAxisVelPrf_Coeff1;
			arAxisVelPrf_Coeff2[iUnitId]:= i_pstStSysParam^.astStUnitParam_Save[iUnitId].rAxisVelPrf_Coeff2;
			arAxisVelPrf_Coeff3[iUnitId]:= i_pstStSysParam^.astStUnitParam_Save[iUnitId].rAxisVelPrf_Coeff3;
		END_FOR
		fbKS_FB_Compensate_Vel_Prn(
			i_xEn:= TRUE,
			i_iGrpId:= i_iGrpId,
			i_rVel_Cur:= i_pstStSysParam^.astStGrpParam_UnSave[i_iGrpId].rVel_Cur,
			i_iGrpUnitNum_Pu:= i_iGrpUnitNum_Pu,
			i_aiGrpUnitList:= i_aiGrpUnitList,
			i_iGrpLinkageAxisNum_Pu:= g_aiGrpLinkageAxisNum_Pu[i_iGrpId],
			i_aiGrpLinkageAxisList:= aiGrpLinkageAxisList,
		//	i_palrAxisMotionVel:= ADR(alrAxisMotionVel),
			i_paxFlag_PressDne:= i_paxFlag_PressDne,
			i_rVel_A:= i_rVel_A,
			i_rVel_Jerk:= i_rVel_Jerk,
			i_arAxisVelPrf_Coeff1:= arAxisVelPrf_Coeff1,//i_pstStSysParam^.astStRSV_GrpParam_Save[i_iGrpId].rAxisVelPrf_Coeff1,
			i_arAxisVelPrf_Coeff2:= arAxisVelPrf_Coeff2,//i_pstStSysParam^.astStRSV_GrpParam_Save[i_iGrpId].rAxisVelPrf_Coeff2,
			i_arAxisVelPrf_Coeff3:= arAxisVelPrf_Coeff3,//i_pstStSysParam^.astStRSV_GrpParam_Save[i_iGrpId].rAxisVelPrf_Coeff3,
			i_xFlag_Accing:= i_pstStSysParam^.astStGrpParam_UnSave[i_iGrpId].xFlag_Accing,
			i_xFlag_Decing:= i_pstStSysParam^.astStGrpParam_UnSave[i_iGrpId].xFlag_Decing,
			o_alrAxisPrfVel=>alrAxisPrfVel);

		FOR iN:=1 TO i_iGrpUnitNum_Pu BY 1 DO
			iUnitId:= i_aiGrpUnitList[iN];
			IF iUnitId>0 AND iUnitId<=MAX_UNIT_NUM THEN
				i_pstStSysParam^.astStUnitParam_UnSave[iUnitId].rAxisPrfVel:= LREAL_TO_REAL(alrAxisPrfVel[iUnitId]);
			END_IF
		END_FOR
//2026.04.11.204941增加结束

		fbKS_FB_AxisVelCtl_PrnRoller(
			i_xEn:= TRUE,
			i_iGrpId:= i_iGrpId,
			i_xSwitchType0:= FALSE,
			i_xSwitchType1:= FALSE,
			i_xMotionStsSwitchEn:= FALSE,
			i_xNeedKeepSync:= FALSE,
			i_iGrpAxisNum_Pu:= i_iGrpUnitNum_Pu,
			i_pstStSysParam:= i_pstStSysParam,
			i_paiGrpAxisList:= ADR(i_aiGrpUnitList),
			i_pastStIOMap_Main_FE:= i_pastStIOMap_Main_FE,
			i_pastStIOMap_Axis_FE:= i_pastStIOMap_Axis_FE,
			i_pabyAxisMotionSts:= ADR(g_abyAxisMotionSts),
			i_paxAxisInching:= ADR(g_axAxisMotionInching),
			i_paxLastAxisInchBtn:= ADR(g_axLastAxisMotionInchBtn),
			i_iMaxVel_StsSwitch:= g_iMaxVel_StsSwitch,
			i_palrAxisMotionVel:= ADR(alrAxisMotionVel),
			i_palrAcceleToSync:= ADR(g_alrAcceleToSync),
			i_palrTimeToSync:= ADR(g_alrTimeToSync),
			i_palrRelatePos_Final:= ADR(g_alrRelatePos_Final),
			i_palrRelatePosToSync:= ADR(g_alrRelatePosToSync),
			i_xMotionEnabled:= i_xMotionEnabled,
			i_xChangLinkageStsWhenPrint:= FALSE,
			i_uiMaxVel_UseCalcAcc:= i_pstStSysParam^.stStSysParam_Save.uiMaxVel_UseCalcAcc,
			o_xEn=> );

		FOR iN:=1 TO  i_iGrpUnitNum_Pu BY 1 DO
			g_alrAxisMotionVel[iN] := alrAxisMotionVel[iN];
		END_FOR

		FOR iN:=1 TO i_iGrpGearMotion_Num BY 1 DO
// 			KS_HY_GetAxisIdForMotByStation(
// 				i_aiGrpGearMotion_StdList[iN],
// 				ADR(iAxisId),
// 				ADR(iTypeId),
// 				ADR(iUnitId),
// 				ADR(iCoreId),
// 				ADR(iGroupId),
// 				ADR(iAdjAxisId),
// 				i_pastStAxisIdListInf);
			KS_GetAxisIdForMotByStation_V2(
					i_iStationId:= i_aiGrpGearMotion_StdList[iN],
					i_piAxisId:= ADR(iAxisId),
					i_piTypeId:= ADR(iTypeId),
					i_piUnitId:= ADR(iUnitId),
					i_piCoreId:= ADR(iCoreId),
					i_piGroupId:= ADR(iGroupId),
					i_piAdjAxisId:= ADR(iAdjAxisId),
					i_pstStSysStationInf:= i_pstStSysStationInf);
			i_pastStMotorParam_Vel^[iN].iAxisId:= iAxisId;
			i_pastStMotorParam_Vel^[iN].iCoreId:= iCoreId;
			i_pastStMotorParam_Vel^[iN].iStationId:= i_aiGrpGearMotion_StdList[iN];
			CASE iTypeId OF
			TYPE_MASTER_I,TYPE_MASTER_II:
				;
			TYPE_CENTRAL_I,TYPE_CENTRAL_II:
				lrTempAxisVel:= pstStGrpParam_UnSave^.rVel_Film;
				IF i_pastStMotorParam_Vel^[iN].xMoveRev THEN
					lrTempAxisVel:= -lrTempAxisVel;
				END_IF
				i_pastStMotorParam_Vel^[iN].rAxisVel:= lrTempAxisVel;
				i_pastStMotorParam_Vel^[iN].rAxisGirth:= pstStGrpParam_Save^.rGirth_CenterRoller;
				i_pastStMotorParam_Vel^[iN].uiAxisNum:= pstStGrpParam_Save^.uiNum_CenterRoller;
				i_pastStMotorParam_Vel^[iN].uiAxisDen:= pstStGrpParam_Save^.uiDen_CenterRoller;
			TYPE_UNWIND_A_I,TYPE_UNWIND_A_II:
				lrTempAxisVel:= pstStGrpParam_UnSave^.rAxisAVelRPM_Cur_Uw;
				IF i_pastStMotorParam_Vel^[iN].xMoveRev THEN
					lrTempAxisVel:= -lrTempAxisVel;
				END_IF
				i_pastStMotorParam_Vel^[iN].rAxisVel:= lrTempAxisVel;
				i_pastStMotorParam_Vel^[iN].uiAxisNum:= pstStGrpParam_Save^.uiNum_Uw;
				i_pastStMotorParam_Vel^[iN].uiAxisDen:= pstStGrpParam_Save^.uiDen_Uw;
			TYPE_UNWIND_B_I,TYPE_UNWIND_B_II:
				lrTempAxisVel:= pstStGrpParam_UnSave^.rAxisBVelRPM_Cur_Uw;
				IF i_pastStMotorParam_Vel^[iN].xMoveRev THEN
					lrTempAxisVel:= -lrTempAxisVel;
				END_IF
				i_pastStMotorParam_Vel^[iN].rAxisVel:= lrTempAxisVel;
				i_pastStMotorParam_Vel^[iN].uiAxisNum:= pstStGrpParam_Save^.uiNum_Uw;
				i_pastStMotorParam_Vel^[iN].uiAxisDen:= pstStGrpParam_Save^.uiDen_Uw;
			TYPE_REWIND_A_I,TYPE_REWIND_A_II:
				lrTempAxisVel:= pstStGrpParam_UnSave^.rAxisAVelRPM_Cur_Rw;
				IF i_pastStMotorParam_Vel^[iN].xMoveRev THEN
					lrTempAxisVel:= -lrTempAxisVel;
				END_IF
				i_pastStMotorParam_Vel^[iN].rAxisVel:= lrTempAxisVel;
				i_pastStMotorParam_Vel^[iN].uiAxisNum:= pstStGrpParam_Save^.uiNum_Rw;
				i_pastStMotorParam_Vel^[iN].uiAxisDen:= pstStGrpParam_Save^.uiDen_Rw;
			TYPE_REWIND_B_I,TYPE_REWIND_B_II:
				lrTempAxisVel:= pstStGrpParam_UnSave^.rAxisBVelRPM_Cur_Rw;
				IF i_pastStMotorParam_Vel^[iN].xMoveRev THEN
					lrTempAxisVel:= -lrTempAxisVel;
				END_IF
				i_pastStMotorParam_Vel^[iN].rAxisVel:= lrTempAxisVel;
				i_pastStMotorParam_Vel^[iN].uiAxisNum:= pstStGrpParam_Save^.uiNum_Rw;
				i_pastStMotorParam_Vel^[iN].uiAxisDen:= pstStGrpParam_Save^.uiDen_Rw;
			TYPE_INFEED_I,TYPE_INFEED_II:
				lrTempAxisVel:= pstStGrpParam_UnSave^.rVel_Cur_If;
				IF i_pastStMotorParam_Vel^[iN].xMoveRev THEN
					lrTempAxisVel:= -lrTempAxisVel;
				END_IF
				i_pastStMotorParam_Vel^[iN].rAxisVel:= lrTempAxisVel;
				i_pastStMotorParam_Vel^[iN].rAxisGirth:= pstStGrpParam_UnSave^.rUsingGirth_If;
				i_pastStMotorParam_Vel^[iN].uiAxisNum:= pstStGrpParam_Save^.uiNum_If;
				i_pastStMotorParam_Vel^[iN].uiAxisDen:= pstStGrpParam_Save^.uiDen_If;
			TYPE_OUTFEED_I,TYPE_OUTFEED_II:
				lrTempAxisVel:= pstStGrpParam_UnSave^.rVel_Cur_Of;
				IF i_pastStMotorParam_Vel^[iN].xMoveRev THEN
					lrTempAxisVel:= -lrTempAxisVel;
				END_IF
				i_pastStMotorParam_Vel^[iN].rAxisVel:= lrTempAxisVel;
				i_pastStMotorParam_Vel^[iN].rAxisGirth:= pstStGrpParam_UnSave^.rUsingGirth_Of;
				i_pastStMotorParam_Vel^[iN].uiAxisNum:= pstStGrpParam_Save^.uiNum_Of;
				i_pastStMotorParam_Vel^[iN].uiAxisDen:= pstStGrpParam_Save^.uiDen_Of;
			TYPE_UNIT_PRN:
				IF pstStGrpParam_UnSave^.xFlag_Stop THEN
					lrTempAxisVel:= i_pstStSysParam^.astStUnitParam_UnSave[iUnitId].rAxisVel_PrnRoller;
				ELSE
					lrTempAxisVel:= alrAxisMotionVel[iUnitId];
				END_IF

				IF i_pastStMotorParam_Vel^[iN].xMoveRev THEN
					lrTempAxisVel:= -lrTempAxisVel;
				END_IF
				i_pastStMotorParam_Vel^[iN].rAxisVel:= lrTempAxisVel;
				i_pastStMotorParam_Vel^[iN].rAxisGirth:= i_pstStSysParam^.astStUnitParam_Save[iUnitId].rGirth_PrnRoller;
				i_pastStMotorParam_Vel^[iN].uiAxisNum:= i_pstStSysParam^.astStUnitParam_Save[iUnitId].uiNum_PrnRoller;
				i_pastStMotorParam_Vel^[iN].uiAxisDen:= i_pstStSysParam^.astStUnitParam_Save[iUnitId].uiDen_PrnRoller;
			TYPE_UNIT_BOTTOM:
				IF g_iMachineryType = MACHINERYTYPE_FELXO_INLINE_ONEBOTOMROLLER THEN //机组式柔印、单伺服底辊
				//	lrTempAxisVel:= alrAxisMotionVel[iUnitId];//i_pstStSysParam^.astStUnitParam_UnSave[iUnitId].rAxisVel_BottomRoller;
					lrTempAxisVel:= i_pstStSysParam^.astStUnitParam_UnSave[iUnitId].rAxisVel_BottomRoller;
				ELSE
					lrTempAxisVel:= i_pstStSysParam^.astStUnitParam_UnSave[iUnitId].rAxisVel_BottomRoller;
				END_IF
				IF i_pastStMotorParam_Vel^[iN].xMoveRev THEN
					lrTempAxisVel:= -lrTempAxisVel;
				END_IF
				i_pastStMotorParam_Vel^[iN].rAxisVel:= lrTempAxisVel;
				i_pastStMotorParam_Vel^[iN].rAxisGirth:= i_pstStSysParam^.astStUnitParam_Save[iUnitId].rGirth_BottomRoller;
				i_pastStMotorParam_Vel^[iN].uiAxisNum:= i_pstStSysParam^.astStUnitParam_Save[iUnitId].uiNum_BottomRoller;
				i_pastStMotorParam_Vel^[iN].uiAxisDen:= i_pstStSysParam^.astStUnitParam_Save[iUnitId].uiDen_BottomRoller;
			TYPE_UNIT_NET:
				lrTempAxisVel:= i_pstStSysParam^.astStUnitParam_UnSave[iUnitId].rAxisVel_NetRoller;
				IF i_pastStMotorParam_Vel^[iN].xMoveRev THEN
					lrTempAxisVel:= -lrTempAxisVel;
				END_IF
				i_pastStMotorParam_Vel^[iN].rAxisVel:= lrTempAxisVel;
				i_pastStMotorParam_Vel^[iN].rAxisGirth:= i_pstStSysParam^.astStUnitParam_Save[iUnitId].rGirth_NetRoller;
				i_pastStMotorParam_Vel^[iN].uiAxisNum:= i_pstStSysParam^.astStUnitParam_Save[iUnitId].uiNum_NetRoller;
				i_pastStMotorParam_Vel^[iN].uiAxisDen:= i_pstStSysParam^.astStUnitParam_Save[iUnitId].uiDen_NetRoller;
			END_CASE
		END_FOR

	i_pastStMotorParam_Vel^[1].rAxisVel;
	i_pastStMotorParam_Vel^[2].rAxisVel;
	i_pastStMotorParam_Vel^[3].rAxisVel;
	i_pastStMotorParam_Vel^[4].rAxisVel;
	i_pastStMotorParam_Vel^[5].rAxisVel;
	i_pastStMotorParam_Vel^[6].rAxisVel;
	i_pastStMotorParam_Vel^[1].xMoveEn;
	i_pastStMotorParam_Vel^[2].xMoveEn;
	i_pastStMotorParam_Vel^[3].xMoveEn;
	i_pastStMotorParam_Vel^[4].xMoveEn;
	i_pastStMotorParam_Vel^[5].xMoveEn;
	i_pastStMotorParam_Vel^[6].xMoveEn;

	END_IF
ELSE
	;
END_IF

(* ---- KS_FB_CheckServeOnDone.st ---- *)
(*@CES
Name=KS_FB_CheckServeOnDone
Type=FunctionBlock
TypeGuid=6f9dac99-8de1-4efc-8465-68ac443b7d08
Guid=4accf54a-639d-49b8-ab4c-ff599b501e0c
HasDeclaration=True
HasImplementation=True
*)
{DECLARATION}
FUNCTION_BLOCK KS_FB_CheckServeOnDone
VAR_INPUT
	i_xEn: BOOL;
	i_iGrpGearMotion_Num: INT;
	i_aiGrpGearMotion_StdList: ARRAY [1..MAX_STATION_NUM] OF INT;
	i_pstStSysParam: POINTER TO StSysParam;
	i_pastStAxisIdListInf :POINTER TO ARRAY [1..128] OF StAxisIdListInf;
	i_pastStGetMotionSts: POINTER TO ARRAY [1..MAX_STATION_NUM] OF StGetMotionSts;
	i_pastStMotorParam_Vel: POINTER TO ARRAY [1..MAX_STATION_NUM] OF StMotorParam_Vel;
	i_xFlag_StopOrEStop : BOOL;
	i_pstStSysStationInf			:POINTER TO StSysStationInf;
END_VAR
VAR_OUTPUT
	o_xEn : BOOL;
	o_xDone : BOOL;
	o_iErrNo : INT;
	o_iErrAxisId : INT;
	o_iErrTypeId : INT;
	o_iErrUnitId : INT;
	o_iErrCoreId : INT;
	o_iErrGroupId : INT;
	o_iErrAdjAxisId : INT;
	o_iMoveErrCode: INT; (* 初始化错误代码
												0-正常
												1-使能异常
												2-模态0设置异常
												3-模态1设置异常
												4-规划器启动异常
												5-PT模式设置异常
												6-伺服打开超时
												7-PT规划异常 *)

END_VAR
VAR
	iN : INT;
	aiErrServoOn_Cnt : ARRAY [1..128] OF INT;
	iServoOnNum : INT;
	iNotNeedServoOnNum : INT;
	iNeedServoOnNum : INT;
	iNeedServoOnNum_Pre : INT;
END_VAR

{IMPLEMENTATION}
o_xEn := i_xEn;
o_iErrNo := 0;
o_iErrAxisId := 0;
o_iErrTypeId := 0;
o_iErrUnitId := 0;
o_iErrCoreId := 0;
iServoOnNum := 0;
iNotNeedServoOnNum := 0;
iNeedServoOnNum := 0;
o_iMoveErrCode := 0;
IF i_xEn THEN
	IF i_pstStSysParam <> 0 AND
		i_pastStAxisIdListInf <> 0 AND
		i_pastStGetMotionSts <> 0 AND
		i_pastStMotorParam_Vel <> 0 AND i_pstStSysStationInf <> 0 THEN
		FOR iN := 1 TO i_iGrpGearMotion_Num BY 1 DO
			IF i_pastStMotorParam_Vel^[iN].xMoveEn THEN
				iNeedServoOnNum := iNeedServoOnNum + 1;
				IF (*i_pastStGetMotionSts^[i_pastStMotorParam_Vel^[iN].iAxisId].dwDriverSts.1 AND*)
					i_pastStGetMotionSts^[i_pastStMotorParam_Vel^[iN].iAxisId].dwMotionSts.9 AND
					//2026.1.20.103746 | + | 运动流程达到写数据的流程
					(i_pastStMotorParam_Vel^[iN].iMoveStep = MOTIONCTL_STEP_WRITEDATA_Run OR
						i_pastStMotorParam_Vel^[iN].iMoveStep = MOTIONCTL_STEP_WRITEDATA_Inch OR
						i_pastStMotorParam_Vel^[iN].iMoveStep = MOTIONCTL_STEP_WRITEDATA_Preg OR
						i_pastStMotorParam_Vel^[iN].iMoveStep = MOTIONCTL_STEP_WRITEDATA_Jog) THEN
					iServoOnNum := iServoOnNum + 1;

					aiErrServoOn_Cnt[iN] := 0;
				ELSE
					aiErrServoOn_Cnt[iN] := aiErrServoOn_Cnt[iN] + 1;
					//2026.1.14.165203 | 伺服等待时间增加到15秒，因为经常出现私服打开超时不知道原因
					IF aiErrServoOn_Cnt[iN] > 15*1000/gc_TENSION_TSK_CYCLE_TIME THEN
						aiErrServoOn_Cnt[iN] := aiErrServoOn_Cnt[iN] -1;
// 						KS_HY_GetAxisIdForMotByStation(
// 							i_aiGrpGearMotion_StdList[iN],
// 							ADR(o_iErrAxisId),
// 							ADR(o_iErrTypeId),
// 							ADR(o_iErrUnitId),
// 							ADR(o_iErrCoreId),
// 							ADR(o_iErrGroupId),
// 							ADR(o_iErrAdjAxisId),
// 							i_pastStAxisIdListInf);
						KS_GetAxisIdForMotByStation_V2(
							i_iStationId:= i_aiGrpGearMotion_StdList[iN],
							i_piAxisId:= ADR(o_iErrAxisId),
							i_piTypeId:= ADR(o_iErrTypeId),
							i_piUnitId:= ADR(o_iErrUnitId),
							i_piCoreId:= ADR(o_iErrCoreId),
							i_piGroupId:= ADR(o_iErrGroupId),
							i_piAdjAxisId:= ADR(o_iErrAdjAxisId),
							i_pstStSysStationInf:= i_pstStSysStationInf);
						o_iMoveErrCode := 6;
						o_iErrNo := -1;
					END_IF
					o_xDone := FALSE;
					EXIT;
				END_IF
			ELSE
				iNotNeedServoOnNum := iNotNeedServoOnNum + 1;
			END_IF
		END_FOR

		IF iServoOnNum = iNeedServoOnNum(*(i_iGrpGearMotion_Num - iNotNeedServoOnNum)*) THEN
			o_xDone := TRUE;
		END_IF
		IF iNeedServoOnNum_Pre <> iNeedServoOnNum THEN
			FOR iN := 1 TO i_iGrpGearMotion_Num BY 1 DO
				aiErrServoOn_Cnt[iN] := 0;
			END_FOR
		END_IF
		iNeedServoOnNum_Pre := iNeedServoOnNum;
	END_IF
ELSE
	IF i_xFlag_StopOrEStop THEN
		o_xDone := FALSE;
	END_IF
END_IF
